(* IEC 61131-3 sources: PLC-IsaVODE/PLC-IsaVODE/samples/plc-programs (part 10) *)

(* ---- 683-FILE_PATH_SPLIT.ST ---- *)
TYPE
  oscat_STRING250             : STRING;
  oscat_STRING1             : STRING;
  oscat_STRING80             : STRING;
  oscat_STRING3             : STRING;
  oscat_NW_BUF_LONG  : ARRAY [0..4095] OF BYTE;
  PRINTF_DATA_250  	:  ARRAY [1..11]  OF oscat_STRING250;
  PRINTF_DATA_80 	:  ARRAY [1..11]  OF oscat_STRING80;
  LOG_250       	:  ARRAY [0..400] OF oscat_STRING250;
  LOG_80    		:  ARRAY [0..400] OF oscat_STRING80;
  LOG_OPTION		:  ARRAY [0..400] OF DWORD;

  us_LOG_CONTROL :
  STRUCT
    NEW_MSG              : oscat_STRING250;    (*W neue Nachricht f�r den Datenbuffer   *)
	NEW_MSG_OPTION 		 : DWORD;
    LEVEL                : BYTE;
	SIZE                 : INT;                (*R Anzahl der Strings im LOG_DATA       *)
	RESET                : BOOL;               (*W Nachrichtenbuffer l�schen            *)
    PRINTF               : PRINTF_DATA_250;    (*W Array PRINTF Parameter               *)
    MSG                  : LOG_250;            (*I Array Message                        *)
    MSG_OPTION           : LOG_OPTION;     	   (*I Array Message Option                 *)
	UPDATE_COUNT         : UINT;               (*R Updatez�hler                         *)
    IDX                  : INT;                (*R aktueller Nachrichten-Index          *)
	RING_MODE            : BOOL;               (*I Buffer�berlauf erkannt               *)
  END_STRUCT;

  us_LOG_CONTROL_80 :
  STRUCT
    NEW_MSG              : oscat_STRING80;     (*W neue Nachricht f�r den Datenbuffer   *)
	NEW_MSG_OPTION 		 : DWORD;
    LEVEL                : BYTE;
	SIZE                 : INT;                (*R Anzahl der Strings im LOG_DATA       *)
	RESET                : BOOL;               (*W Nachrichtenbuffer l�schen            *)
    PRINTF               : PRINTF_DATA_80;     (*W Array PRINTF Parameter               *)
    MSG                  : LOG_80;             (*I Array Message                        *)
    MSG_OPTION           : LOG_OPTION;     	   (*I Array Message Option                 *)
	UPDATE_COUNT         : UINT;               (*R Updatez�hler                         *)
    IDX                  : INT;                (*R aktueller Nachrichten-Index          *)
	RING_MODE            : BOOL;               (*I Buffer�berlauf erkannt               *)
  END_STRUCT;

  LINE_ARRAY 			: ARRAY [1..40] OF INT;

  us_LOG_VIEWPORT :
    STRUCT
     LINE_ARRAY          : LINE_ARRAY;
     COUNT               : INT;                (* Anzahl der sichtbaren Nachtrichten   *)
	 UPDATE_COUNT        : UINT;               (* Updatez�hler                         *)
     MOVE_TO_X           : INT;                (* Steuerung der Nachrichtenanzeige     *)
     UPDATE              : BOOL;               (* Daten wurden ge�ndert -> neuzeichnen *)
  END_STRUCT;

  oscat_FILE_SERVER_DATA : STRUCT
	FILE_OPEN	: BOOL;
    FILENAME 	: STRING;
    MODE	 	: BYTE;
    OFFSET   	: UDINT;
    FILE_SIZE   : UDINT;
    AUTO_CLOSE	: TIME;
    ERROR	 	: BYTE;
  END_STRUCT;

  oscat_FILE_PATH_DATA : STRUCT
	DRIVE : oscat_string3;
	DIRECTORY : oscat_string250;
	FILENAME : STRING;
  END_STRUCT;

  oscat_UNI_CIRCULAR_BUFFER_DATA : STRUCT
	D_MODE : INT;
	D_HEAD : WORD;
	D_STRING : oscat_string250;
	D_REAL : REAL;
	D_DWORD : DWORD;
	BUF_SIZE : INT;
	BUF_COUNT : INT;
	BUF_USED : USINT;
	BUF : oscat_NW_BUF_LONG;
	_GetStart : INT;
	_GetEnd : INT;
	_Last : INT;
	_First : INT;
  END_STRUCT;

  oscat_DLOG_DATA : STRUCT
	STORE_TYPE : BYTE;
	ADD_HEADER : BOOL;
	ADD_DATA : BOOL;
	ADD_DATA_REQ : BOOL;
	CLOCK_TRIG : BOOL;
	ID_MAX : USINT;
	DTI : UDINT;
	UCB : oscat_UNI_CIRCULAR_BUFFER_DATA;
	NEW_FILE : STRING;
	NEW_FILE_RTRIG : BOOL;
  END_STRUCT;

END_TYPE

FUNCTION_BLOCK FILE_PATH_SPLIT_Block

	VAR_INPUT
		FILENAME :	oscat_STRING250;
	END_VAR

	VAR_OUTPUT
		FILE_PATH_SPLIT :	BOOL;
	END_VAR

	VAR_IN_OUT
		X :	oscat_FILE_PATH_DATA;
	END_VAR

	VAR
		b :	INT;
		c :	INT;
		d :	oscat_STRING1;
		p1 :	INT;
		p2 :	INT;
	END_VAR

	X.DRIVE := '';
	X.DIRECTORY := '';
	X.FILENAME := '';
	p1 := 0;
	p2 := 0;
	c := LEN(FILENAME);
	IF c = 0 THEN
		FILE_PATH_SPLIT := FALSE;
		RETURN;
	END_IF;

	FOR b := 1 TO c DO
		d := MID(FILENAME, 1, b);
		IF EQ_STRING(d,':') THEN
			p1 := b;
		ELSIF EQ_STRING(d,'/') OR EQ_STRING(d,'\') THEN
			p2 := b;
		END_IF;
	END_FOR;

	IF p1 = 2 THEN
		X.DRIVE := LEFT(FILENAME,p1);
	END_IF;

	IF p2 > 0 AND p2 > p1 THEN
		X.DIRECTORY := MID(FILENAME,p2-p1,p1+1);
	END_IF;

	X.FILENAME := RIGHT(FILENAME,c - MAX (p1,p2));
	FILE_PATH_SPLIT := TRUE;

END_FUNCTION_BLOCK

PROGRAM program0
	VAR
		FILENAME :	oscat_STRING250;
		FILE_PATH_SPLIT :	BOOL;
		X :	oscat_FILE_PATH_DATA;

		func_block : FILE_PATH_SPLIT_Block;
	END_VAR
	func_block.FILENAME := FILENAME;
	func_block.X := X;

	func_block();
	FILE_PATH_SPLIT  := func_block.FILE_PATH_SPLIT;
	X  := func_block.X;
END_PROGRAM

CONFIGURATION Config0
	RESOURCE Res0 ON PLC
		TASK task0(INTERVAL := T#20ms,PRIORITY := 0);
		PROGRAM instance0 WITH task0 : program0;
	END_RESOURCE
END_CONFIGURATION

(* ---- 684-BLIND_SHADE.ST ---- *)
TYPE
  oscat_STRING5               : STRING;
  oscat_STRING30              : STRING;
END_TYPE

TYPE oscat_CALENDAR :
	STRUCT
		UTC : UDINT;				(* world time UTC *)
		LDT : UDINT;				(* local time *)
		LDATE : UDINT;				(* local date *)
		LTOD : UDINT;				(* local time of day *)
		YEAR : INT;					(* year of LDATE *)
		MONTH : INT;				(* month of LDATE *)
		DAY : INT;					(* day of LDATE *)
		WEEKDAY : INT;				(* weekday of LDATE *)
		OFFSET : INT;				(* Time Zone Offset for Local time in minutes *)
		DST_EN : BOOL;				(* daylight savings time enable *)
		DST_ON : BOOL;				(* true when daylight savings time os on *)
		NAME : oscat_string5;		(* name of time zone *)
		LANGUAGE : INT;			    (* language number pls see language setup *)
		LONGITUDE : REAL;			(* longitude of current location *)
		LATITUDE : REAL;			(* latitude of current location *)
		SUN_RISE : UDINT;			(* sun_rise for current location *)
		SUN_SET : UDINT;			(* sun_set for current location *)
		SUN_MIDDAY : UDINT;			(* worldtime when sun stands at south position *)
		SUN_HEIGTH : REAL;			(* suns heigth at midday, south position *)
		SUN_HOR : REAL;				(* sun angle horizontal 0 = north in degrees *)
		SUN_VER : REAL;				(* sun angle vertical above horizon in degrees *)
		NIGHT : BOOL;				(* true between sun_set and sun_rise *)
		HOLIDAY : BOOL;				(* true when holiday *)
		HOLY_NAME : oscat_string30;	(* name of holiday *)
		WORK_WEEK : INT;			(* current work week *)
	END_STRUCT;
END_TYPE

FUNCTION DT_TO_TOD2:UDINT
	VAR_INPUT
		IN :	UDINT;
	END_VAR

	DT_TO_TOD2 := (IN MOD UDINT#86400) * UDINT#1000;
END_FUNCTION

FUNCTION TIME_TO_UDINT2:UDINT
	VAR_INPUT
		X :	TIME;
	END_VAR

	TIME_TO_UDINT2 := DINT_TO_UDINT(TIME_TO_DINT(X));
END_FUNCTION

FUNCTION DEG : REAL
	VAR_INPUT
		RAD_IN : REAL;
	END_VAR

	DEG := MODR(57.29577951308232 * RAD_IN, 360.0);
END_FUNCTION

FUNCTION MODR : REAL
	VAR_INPUT
		IN : REAL;
		DIVI : REAL;
	END_VAR

	IF divi = 0.0 THEN
		MODR := 0.0;
	ELSE
		MODR := in - DINT_TO_REAL(FLOOR2(in / divi)) * divi;
	END_IF;
END_FUNCTION

FUNCTION FLOOR2 : DINT
	VAR_INPUT
		x : REAL;
	END_VAR

	FLOOR2 := REAL_TO_DINT(X);
	IF DINT_TO_REAL(FLOOR2) > X THEN
		FLOOR2 := FLOOR2 - DINT#1;
	END_IF;
END_FUNCTION

FUNCTION RAD:REAL

	VAR_INPUT
		DEG1 :	REAL;
	END_VAR

	RAD := MODR(0.0174532925199433 * DEG1 , 6.283185307179586476);

END_FUNCTION

FUNCTION TRUNC_UDINT2:UDINT
	VAR_INPUT
		IN :	REAL;
	END_VAR
	TRUNC_UDINT2 := DINT_TO_UDINT(TRUNC_DINT(IN));
END_FUNCTION

FUNCTION_BLOCK BLIND_SHADE_Block

	VAR_INPUT
		UP :	BOOL;
		DN :	BOOL;
		S_IN :	BYTE;
		PI :	BYTE;
		AI :	BYTE;
		ENABLE :	BOOL;
		SUN :	BOOL;
		SUNRISE_OFFSET :	TIME := T#1h;
		SUNSET_PRESET :	TIME := T#1h;
		DIRECTION :	REAL := 180.0;
		ANGLE_OFFSET :	REAL := 80.0;
		SLAT_WIDTH :	REAL := 80.0;
		SLAT_SPACING :	REAL := 60.0;
		SHADE_DELAY :	TIME := T#60s;
		SHADE_POS :	BYTE;
	END_VAR

	VAR_OUTPUT
		QU :	BOOL;
		QD :	BOOL;
		STATUS :	BYTE;
		PO :	BYTE;
		AO :	BYTE;
	END_VAR

	VAR_IN_OUT
		CX :	oscat_CALENDAR;
	END_VAR

	VAR
		angle :	REAL;
		sun_delay :	TOF;
	END_VAR

	sun_delay(IN := sun, PT := shade_delay);

	IF UP AND DN AND enable AND sun_delay.Q AND cx.SUN_HOR > direction - angle_offset AND cx.SUN_HOR < direction + angle_offset AND
		DT_TO_TOD2(cx.UTC) > cx.SUN_RISE + TIME_TO_UDINT2(sunrise_offset) AND DT_TO_TOD2(cx.UTC) < cx.SUN_SET - TIME_TO_UDINT2(sunset_preset) THEN
		status := BYTE#151;
		QU := UP;
		QD := DN;
		po := shade_pos;
		angle := DEG(ATAN(slat_spacing / slat_width));
		IF cx.SUN_VER > 0.0 AND cx.SUN_VER < angle THEN
			angle := cx.SUN_VER + DEG(ACOS(COS(RAD(cx.SUN_VER))*slat_spacing / Slat_width));
			ao := INT_TO_BYTE(LIMIT(0,UDINT_TO_INT(TRUNC_UDINT2(angle * 2.833333333)), 255));
		ELSE
			ao := BYTE#255;
		END_IF;
	ELSE
		QU := UP;
		QD := DN;
		po := pi;
		ao := ai;
		status := S_IN;
	END_IF;

END_FUNCTION_BLOCK

PROGRAM program0
	VAR
		UP :	BOOL;
		DN :	BOOL;
		S_IN :	BYTE;
		PI :	BYTE;
		AI :	BYTE;
		ENABLE :	BOOL;
		SUN :	BOOL;
		SUNRISE_OFFSET :	TIME := T#1h;
		SUNSET_PRESET :	TIME := T#1h;
		DIRECTION :	REAL := 180.0;
		ANGLE_OFFSET :	REAL := 80.0;
		SLAT_WIDTH :	REAL := 80.0;
		SLAT_SPACING :	REAL := 60.0;
		SHADE_DELAY :	TIME := T#60s;
		SHADE_POS :	BYTE;
		CX :	oscat_CALENDAR;

		func_block : BLIND_SHADE_Block;
	END_VAR
	func_block.UP := UP;
	func_block.DN := DN;
	func_block.S_IN := S_IN ;
	func_block.PI    := PI    ;
	func_block.AI    := AI    ;
	func_block.ENABLE := ENABLE;
	func_block.SUN := SUN;
	func_block.SUNRISE_OFFSET := SUNRISE_OFFSET;
	func_block.SUNSET_PRESET := SUNSET_PRESET ;
	func_block.DIRECTION := DIRECTION ;
	func_block.ANGLE_OFFSET    := ANGLE_OFFSET    ;
	func_block.SLAT_WIDTH := SLAT_WIDTH;
	func_block.SLAT_SPACING := SLAT_SPACING;
	func_block.SHADE_DELAY := SHADE_DELAY ;
	func_block.CX := CX ;

	func_block();
	CX  := func_block.CX;
END_PROGRAM

CONFIGURATION Config0
	RESOURCE Res0 ON PLC
		TASK task0(INTERVAL := T#20ms,PRIORITY := 0);
		PROGRAM instance0 WITH task0 : program0;
	END_RESOURCE
END_CONFIGURATION

(* ---- 686-_ARRAY_SHUFFLE.ST ---- *)
TYPE
	oscat_pt_ARRAY: ARRAY [1..100] OF REAL;
END_TYPE

FUNCTION D_TRUNC : DINT
  VAR_INPUT
    x : REAL;
  END_VAR

  D_TRUNC := REAL_TO_DINT(X);
  IF X > 0.0 THEN
  	IF DINT_TO_REAL(D_TRUNC) > X THEN D_TRUNC := D_TRUNC - DINT#1; END_IF;
  ELSE
  	IF DINT_TO_REAL(D_TRUNC) < X THEN D_TRUNC := D_TRUNC + DINT#1; END_IF;
  END_IF;
END_FUNCTION

FUNCTION BIT_COUNT:INT
	VAR_INPUT
		IN :	DWORD;
	END_VAR

	VAR
		in_temp :	DWORD;
	END_VAR

	in_temp := IN;
	WHILE in_temp > DWORD#0 DO
		IF (in_temp AND DWORD#16#00000001) > DWORD#0 THEN Bit_Count := Bit_Count +1; END_IF;
		in_temp := SHR(in_temp,1);
	END_WHILE;
END_FUNCTION

FUNCTION FRACT:REAL
	VAR_INPUT
		X :	REAL;
	END_VAR

	IF ABS(x) < 2.0E9 THEN
		FRACT := x - DINT_TO_REAL(D_TRUNC(x));
	ELSE
		FRACT := 0.0;
	END_IF;
END_FUNCTION

FUNCTION_BLOCK T_PLC_MS_block
	VAR_OUTPUT
		T_PLC_MS :	UDINT;
	END_VAR

	VAR_EXTERNAL
		PLC_TICKS_PER_SEC :	INT;
		PLC_SYS_TICK_CNT :	DINT;
	END_VAR

	VAR
		debug :	BOOL;(*Debug-Mode ON / OFF*)
		N :	INT;(*Debug-Faktor*)
		Offset :	UDINT;(*Debug-Offset*)
		temp :	DWORD := DWORD#1;(*Debug-Offset*)
		mode :	BOOL;(*modus*)
		faktor :	UDINT;(*Systemtakt-Faktor*)
		init :	BOOL;
		v_plc_ticks_per_sec :	UDINT;
		base :	UDINT := UDINT#1000;
	END_VAR

	IF init = FALSE THEN
		v_plc_ticks_per_sec := INT_TO_UDINT(PLC_TICKS_PER_SEC);
		IF v_plc_ticks_per_sec = UDINT#1024 THEN
			faktor := UDINT#1;
			mode := FALSE;
		ELSIF v_plc_ticks_per_sec > UDINT#0 THEN
			IF v_plc_ticks_per_sec <= base THEN
				faktor := base / v_plc_ticks_per_sec;
				mode := FALSE;
			ELSE
				faktor := v_plc_ticks_per_sec / base;
				mode := TRUE;
			END_IF;
		ELSE
			faktor := UDINT#1;
		END_IF;
		init := TRUE;
	END_IF;

	IF mode THEN
		T_PLC_MS := DINT_TO_UDINT(PLC_SYS_TICK_CNT) / faktor;
	ELSE
		T_PLC_MS := DINT_TO_UDINT(PLC_SYS_TICK_CNT) * faktor;
	END_IF;

	IF debug THEN
		T_PLC_MS := (DWORD_TO_UDINT(SHL(UDINT_TO_DWORD(T_PLC_MS),N) OR SHL(temp,N)) - UDINT#1) + Offset;
	END_IF;
END_FUNCTION_BLOCK

FUNCTION BIT_LOAD_DW:DWORD

	VAR_INPUT
		IN :	DWORD;
		VAL :	BOOL;
		POS :	INT;
	END_VAR

	IF val THEN
		BIT_LOAD_DW := in OR SHL(DWORD#1,pos);
	ELSE
		BIT_LOAD_DW := in AND (NOT SHL(DWORD#1,pos));
	END_IF;
END_FUNCTION

FUNCTION BIT_OF_DWORD : BOOL
  VAR_INPUT
    IN : DWORD;
    N : INT;
  END_VAR

  BIT_OF_DWORD := (SHR(in,N) AND 16#00000001) > 0;
  (* from OSCAT library; www.oscat.de  *)
END_FUNCTION

FUNCTION _INT_TO_UDINT:UDINT
	VAR_INPUT
		IN :	INT;
	END_VAR

	_INT_TO_UDINT := DINT_TO_UDINT(INT_TO_DINT(IN));
END_FUNCTION

FUNCTION _DWORD_TO_REAL:REAL
	VAR_INPUT
		IN :	DWORD;
	END_VAR

	_DWORD_TO_REAL := UDINT_TO_REAL(DWORD_TO_UDINT(IN));

END_FUNCTION

FUNCTION_BLOCK RDM_block
	VAR_INPUT
		LAST :	REAL;
	END_VAR
	VAR_OUTPUT
		RDM :	REAL;
	END_VAR
	VAR
		T_PLC_MS :	T_PLC_MS_block;
		tn :	DWORD;
		tc :	INT;
	END_VAR
	T_PLC_MS();
	tn := UDINT_TO_DWORD(T_PLC_MS.T_PLC_MS);
	tc := Bit_Count(tn);

	tn:=BIT_LOAD_DW(tn,BIT_OF_DWORD(tn,2),31); (* tn.31 := tn.2; *)
	tn:=BIT_LOAD_DW(tn,BIT_OF_DWORD(tn,5),30); (* tn.30 := tn.5; *)
	tn:=BIT_LOAD_DW(tn,BIT_OF_DWORD(tn,4),29); (* tn.29 := tn.4; *)
	tn:=BIT_LOAD_DW(tn,BIT_OF_DWORD(tn,1),28); (* tn.28 := tn.1; *)
	tn:=BIT_LOAD_DW(tn,BIT_OF_DWORD(tn,0),27); (* tn.27 := tn.0; *)
	tn:=BIT_LOAD_DW(tn,BIT_OF_DWORD(tn,7),26); (* tn.26 := tn.7; *)
	tn:=BIT_LOAD_DW(tn,BIT_OF_DWORD(tn,6),25); (* tn.25 := tn.6; *)
	tn:=BIT_LOAD_DW(tn,BIT_OF_DWORD(tn,3),24); (* tn.24 := tn.3; *)

	tn := ROL(tn,Bit_Count(tn)) OR DWORD#16#80000001;
	tn := UDINT_TO_DWORD(DWORD_TO_UDINT(tn) MOD UDINT#71474513 + _INT_TO_UDINT(tc) + UDINT#77);
	RDM := fract(_DWORD_TO_REAL(tn) / 10000000.0 * (2.71828182845904523536028747135266249 - LIMIT_REAL(0.0,last,1.0)));
END_FUNCTION_BLOCK

FUNCTION_BLOCK RDM22
	VAR_INPUT
		LAST :	INT;
		LOW :	INT;
		HIGH :	INT;
	END_VAR

	VAR_OUTPUT
		RDM2 :	INT;
	END_VAR

	VAR
		rdm :	RDM_block;
	END_VAR

	rdm(last:=fract(INT_TO_REAL(last) * 3.14159265358979323846264338327950288));
	RDM2 := TRUNC(rdm.RDM * INT_TO_REAL(high - low + 1)) + low;
END_FUNCTION_BLOCK

FUNCTION_BLOCK _ARRAY_SHUFFLE2
	VAR_IN_OUT
		PT :	oscat_pt_ARRAY;
	END_VAR

	VAR_INPUT
		SIZE :	UINT;
	END_VAR

	VAR_OUTPUT
		_ARRAY_SHUFFLE :	BOOL;
	END_VAR
	VAR
		temp :	REAL;
		pos :	INT;
		i :	INT;
		stop :	INT;
		rdm2 :	rdm22;
	END_VAR

	stop :=LIMIT_INT(1,UINT_TO_INT(size),1000);
	FOR i := 1 TO stop DO
			rdm2(last:=i+pos,low:=1,high:=stop);
			pos := rdm2.rdm2;
			(* swap elements *)
			temp := pt[i];
			pt[i] := pt[pos];
			pt[pos] := temp;
	END_FOR;

	_ARRAY_SHUFFLE := TRUE;
END_FUNCTION_BLOCK

PROGRAM program0
  VAR
    LocalVar0 : oscat_pt_ARRAY;
    LocalVar1 : UINT;
	LocalOUT  : BOOL;
	func_block : _ARRAY_SHUFFLE2;
  END_VAR
	func_block.pt := LocalVar0;
	func_block.size := LocalVar1;
	func_block();
	LocalOUT := func_block._ARRAY_SHUFFLE;

END_PROGRAM

CONFIGURATION Config0
	VAR_GLOBAL
		PLC_TICKS_PER_SEC :	INT;
		PLC_SYS_TICK_CNT :	DINT;
	END_VAR
  RESOURCE Res0 ON PLC
    TASK task0(INTERVAL := T#20ms,PRIORITY := 0);
    PROGRAM instance0 WITH task0 : program0;
  END_RESOURCE
END_CONFIGURATION

(* ---- 687-TN_INPUT_SELECT_TEXT.ST ---- *)
TYPE
  bya_TN_CHAR:       	ARRAY [0..1919] OF BYTE;
  bya_TN_BACKUP:     	ARRAY [0..1919] OF BYTE;
  bya_TN_COLOR:      	ARRAY [0..1919] OF BYTE;
  bya_TN_Line_Update:	ARRAY [0..23]   OF BOOL;

  us_TN_SCREEN :
  STRUCT
		bya_CHAR:			bya_TN_CHAR;
		bya_COLOR:			bya_TN_COLOR;
		bya_BACKUP:			bya_TN_BACKUP;
		bya_Line_Update:	bya_TN_Line_Update;

		by_Input_Exten_Code:    BYTE;
		by_Input_ASCII_Code:    BYTE;
		bo_Input_ASCII_IsNum:   BOOL;
		in_Page_Number:        	INT;
		in_Cursor_X:           	INT;
		in_Cursor_Y:           	INT;
		in_EOS_Offset:         	INT;
		by_Clear_Screen_Attr:  	BYTE;
		bo_Clear_Screen:       	BOOL;
		bo_Modal_Dialog:       	BOOL;
		bo_Menue_Bar_Dialog:   	BOOL;

  END_STRUCT;
END_TYPE

FUNCTION_BLOCK TN_INPUT_SELECT_TEXT_Block

  VAR
    in_count :	INT;
    by_Attr :	BYTE;
    st_String :	STRING;
  END_VAR

  VAR
    FB_FIX :	FIX;
    FB_TN_SC_WRITE :	TN_SC_WRITE;
    ELEMENT_COUNT :	ELEMENT_COUNT;
    ELEMENT_GET :	ELEMENT_GET;
  END_VAR

  VAR_IN_OUT
    Xus_TN_SCREEN :	us_TN_SCREEN;
    Xus_TN_INPUT_CONTROL_DATA :	us_TN_INPUT_CONTROL_DATA;
  END_VAR

  IF Xus_TN_INPUT_CONTROL_DATA.bo_Focus = TRUE THEN

    IF Xus_TN_INPUT_CONTROL_DATA.by_Input_ASCII_Code = BYTE#32 THEN
      Xus_TN_INPUT_CONTROL_DATA.in_selected := Xus_TN_INPUT_CONTROL_DATA.in_selected + INT#01;
      Xus_TN_INPUT_CONTROL_DATA.bo_Update_Input := TRUE;
    END_IF;

    IF Xus_TN_INPUT_CONTROL_DATA.by_Input_Exten_Code = BYTE#13 THEN
      Xus_TN_INPUT_CONTROL_DATA.bo_Input_Entered := TRUE;
    END_IF;

  END_IF;

  IF (Xus_TN_INPUT_CONTROL_DATA.bo_Update_Input = TRUE) OR (Xus_TN_INPUT_CONTROL_DATA.bo_Update_All = TRUE) THEN

    IF Xus_TN_INPUT_CONTROL_DATA.bo_Update_All = TRUE THEN

      IF (Xus_TN_INPUT_CONTROL_DATA.in_Title_X_Offset = INT#00) AND (Xus_TN_INPUT_CONTROL_DATA.in_Title_Y_Offset = INT#00) THEN

        FB_TN_SC_WRITE.Iin_Y := Xus_TN_INPUT_CONTROL_DATA.in_Y;
        FB_TN_SC_WRITE.Iin_X := Xus_TN_INPUT_CONTROL_DATA.in_X - LEN(Xus_TN_INPUT_CONTROL_DATA.st_Title_String);

      ELSE
        FB_TN_SC_WRITE.Iin_Y := Xus_TN_INPUT_CONTROL_DATA.in_Y + Xus_TN_INPUT_CONTROL_DATA.in_Title_Y_Offset;
        FB_TN_SC_WRITE.Iin_X := Xus_TN_INPUT_CONTROL_DATA.in_X + Xus_TN_INPUT_CONTROL_DATA.in_Title_X_Offset;

      END_IF;

      FB_TN_SC_WRITE.Iby_ATTR      := Xus_TN_INPUT_CONTROL_DATA.by_Title_Attr;
      FB_TN_SC_WRITE.Ist_STRING    := Xus_TN_INPUT_CONTROL_DATA.st_Title_String;
      FB_TN_SC_WRITE.Xus_TN_SCREEN := Xus_TN_SCREEN;
      FB_TN_SC_WRITE();
      Xus_TN_SCREEN := FB_TN_SC_WRITE.Xus_TN_SCREEN;

    END_IF;

    ELEMENT_COUNT(ELEMENT:=Xus_TN_INPUT_CONTROL_DATA.st_Input_Data,SEP:=BYTE#35);
    Xus_TN_INPUT_CONTROL_DATA.st_Input_Data:=ELEMENT_COUNT.ELEMENT;
    in_count:=ELEMENT_COUNT.ELEMENT_COUNT;

    IF in_Count > INT#00 THEN

      IF Xus_TN_INPUT_CONTROL_DATA.in_selected < INT#1 THEN
        Xus_TN_INPUT_CONTROL_DATA.in_selected := INT#01;
      END_IF;

      IF Xus_TN_INPUT_CONTROL_DATA.in_selected > in_count THEN
        Xus_TN_INPUT_CONTROL_DATA.in_selected := INT#01;
      END_IF;

      ELEMENT_GET(ELEMENT:=Xus_TN_INPUT_CONTROL_DATA.st_Input_Data,SEP:=BYTE#35,POS:=Xus_TN_INPUT_CONTROL_DATA.in_selected-1);
      Xus_TN_INPUT_CONTROL_DATA.st_Input_Data := ELEMENT_GET.ELEMENT;
      st_String:=ELEMENT_GET.ELEMENT_GET;

      FB_FIX.str:=st_String;
    FB_FIX.L:=LEN(Xus_TN_INPUT_CONTROL_DATA.st_Input_Mask);
    FB_FIX.C:=BYTE#32;
    FB_FIX.M:=Xus_TN_INPUT_CONTROL_DATA.in_Input_Option;
      FB_FIX();
      st_String:=FB_FIX.FIX;

      Xus_TN_INPUT_CONTROL_DATA.st_Input_String := st_String;

      IF Xus_TN_INPUT_CONTROL_DATA.bo_Focus = TRUE THEN
        by_Attr := Xus_TN_INPUT_CONTROL_DATA.by_Attr_mF;
      ELSE
        by_Attr := Xus_TN_INPUT_CONTROL_DATA.by_Attr_oF;
      END_IF;

      FB_TN_SC_WRITE.Iin_Y         := Xus_TN_INPUT_CONTROL_DATA.in_Y;
      FB_TN_SC_WRITE.Iin_X         := Xus_TN_INPUT_CONTROL_DATA.in_X;
      FB_TN_SC_WRITE.Iby_ATTR      := by_Attr;
      FB_TN_SC_WRITE.Ist_STRING    := st_String;
      FB_TN_SC_WRITE.Xus_TN_SCREEN := Xus_TN_SCREEN;
      FB_TN_SC_WRITE();
      Xus_TN_SCREEN := FB_TN_SC_WRITE.Xus_TN_SCREEN;

    END_IF;

    Xus_TN_INPUT_CONTROL_DATA.in_Cursor_Y := Xus_TN_INPUT_CONTROL_DATA.in_Y;
    Xus_TN_INPUT_CONTROL_DATA.in_Cursor_X := Xus_TN_INPUT_CONTROL_DATA.in_X;

    Xus_TN_INPUT_CONTROL_DATA.bo_Update_All   := FALSE;
    Xus_TN_INPUT_CONTROL_DATA.bo_Update_Input := FALSE;

  END_IF;

END_FUNCTION_BLOCK

PROGRAM program0
	VAR
		Xus_TN_SCREEN :	us_TN_SCREEN;
    Xus_TN_INPUT_CONTROL_DATA :	us_TN_INPUT_CONTROL_DATA;

		func_block : TN_INPUT_SELECT_TEXT_Block;
	END_VAR
	func_block.Xus_TN_INPUT_CONTROL_DATA := Xus_TN_INPUT_CONTROL_DATA;
	func_block.Xus_TN_SCREEN := Xus_TN_SCREEN;

	func_block();
  Xus_TN_INPUT_CONTROL_DATA  := func_block.Xus_TN_INPUT_CONTROL_DATA;
	Xus_TN_SCREEN  := func_block.Xus_TN_SCREEN;
END_PROGRAM

CONFIGURATION Config0
	RESOURCE Res0 ON PLC
		TASK task0(INTERVAL := T#20ms,PRIORITY := 0);
		PROGRAM instance0 WITH task0 : program0;
	END_RESOURCE
END_CONFIGURATION

(* ---- 688-SEQUENCE_4.ST ---- *)
FUNCTION UDINT_TO_TIME2:TIME

	VAR_INPUT
		IN :	UDINT;
	END_VAR

	UDINT_TO_TIME2 := DINT_TO_TIME(UDINT_TO_DINT(IN));

END_FUNCTION

FUNCTION_BLOCK T_PLC_MS_block
	VAR_OUTPUT
		T_PLC_MS :	UDINT;
	END_VAR

	VAR_EXTERNAL
		PLC_TICKS_PER_SEC :	INT;
		PLC_SYS_TICK_CNT :	DINT;
	END_VAR

	VAR
		debug :	BOOL;
		N :	INT;
		Offset :	UDINT;
		temp :	DWORD := DWORD#1;
		mode :	BOOL;
		faktor :	UDINT;
		init :	BOOL;
		v_plc_ticks_per_sec :	UDINT;
		base :	UDINT := UDINT#1000;
	END_VAR

	IF init = FALSE THEN
		v_plc_ticks_per_sec := INT_TO_UDINT(PLC_TICKS_PER_SEC);
		IF v_plc_ticks_per_sec = UDINT#1024 THEN
			faktor := UDINT#1;
			mode := FALSE;
		ELSIF v_plc_ticks_per_sec > UDINT#0 THEN
			IF v_plc_ticks_per_sec <= base THEN
				faktor := base / v_plc_ticks_per_sec;
				mode := FALSE;
			ELSE
				faktor := v_plc_ticks_per_sec / base;
				mode := TRUE;
			END_IF;
		ELSE
			faktor := UDINT#1;
		END_IF;
		init := TRUE;
	END_IF;

	IF mode THEN
		T_PLC_MS := DINT_TO_UDINT(PLC_SYS_TICK_CNT) / faktor;
	ELSE
		T_PLC_MS := DINT_TO_UDINT(PLC_SYS_TICK_CNT) * faktor;
	END_IF;

	IF debug THEN
		T_PLC_MS := (DWORD_TO_UDINT(SHL(UDINT_TO_DWORD(T_PLC_MS),N) OR SHL(temp,N)) - UDINT#1) + Offset;
	END_IF;

END_FUNCTION_BLOCK

FUNCTION_BLOCK SEQUENCE_4_Block

	VAR_INPUT
		IN0 :	BOOL := TRUE;
		IN1 :	BOOL := TRUE;
		IN2 :	BOOL := TRUE;
		IN3 :	BOOL := TRUE;
		START :	BOOL;
		RST :	BOOL;
		WAIT0 :	TIME;
		DELAY0 :	TIME;
		WAIT1 :	TIME;
		DELAY1 :	TIME;
		WAIT2 :	TIME;
		DELAY2 :	TIME;
		WAIT3 :	TIME;
		DELAY3 :	TIME;
		STOP_ON_ERROR :	BOOL;
	END_VAR

	VAR_OUTPUT
		Q0 :	BOOL;
		Q1 :	BOOL;
		Q2 :	BOOL;
		Q3 :	BOOL;
		QX :	BOOL;
		RUN :	BOOL;
		_STEP :	INT := -1;
		STATUS :	BYTE;
	END_VAR

	VAR
		last :	TIME;
		edge :	BOOL;
		tx :	TIME;
		init :	BOOL;
		T_PLC_MS :	T_PLC_MS_Block;
	END_VAR

	T_PLC_MS();
	tx:= UDINT_TO_TIME(T_PLC_MS.T_PLC_MS);

	IF NOT init THEN
		last := tx;
		init := TRUE;
		status := BYTE#110;
	END_IF;

	IF rst THEN
		_step := -1;
		Q0 := FALSE;
		Q1 := FALSE;
		Q2 := FALSE;
		Q3 := FALSE;
		status := BYTE#110;
		run := FALSE;

	ELSIF start AND NOT edge THEN
		_step := 0;
		last := tx;
		status := BYTE#111;
		Q0 := FALSE;
		Q1 := FALSE;
		Q2 := FALSE;
		Q3 := FALSE;
		run := TRUE;
	END_IF;
	edge := start;

	IF status > BYTE#0 AND status < BYTE#100 AND stop_on_error THEN RETURN; END_IF;

	IF run AND _step = 0 THEN
		IF NOT q0 AND in0 AND tx - last <= wait0 THEN
			Q0 := TRUE;
			last := tx;
		ELSIF NOT q0 AND tx - last > wait0 THEN
			status := BYTE#1;
			run := FALSE;
		ELSIF q0 AND tx - last >= delay0 THEN
			_step := 1;
			last := tx;
		END_IF;
	END_IF;
	IF run AND _step = 1 THEN
		IF NOT q1 AND in1 AND tx - last <= wait1 THEN
			Q0 := FALSE;
			Q1 := TRUE;
			last := tx;
		ELSIF NOT q1 AND Tx - last > wait1 THEN
			status := BYTE#2;
			q0 := FALSE;
			run := FALSE;
		ELSIF q1 AND tx - last >= delay1 THEN
			_step := 2;
			last := tx;
		END_IF;
	END_IF;
	IF run AND _step = 2 THEN
		IF NOT q2 AND in2 AND tx - last <= wait2 THEN
			Q1 := FALSE;
			Q2 := TRUE;
			last := tx;
		ELSIF NOT q2 AND Tx - last > wait2 THEN
			status := BYTE#3;
			q1 := FALSE;
			run := FALSE;
		ELSIF q2 AND tx - last >= delay2 THEN
			_step := 3;
			last := tx;
		END_IF;
	END_IF;
	IF run AND _step = 3 THEN
		IF NOT q3 AND in3 AND tx - last <= wait3 THEN
			Q2 := FALSE;
			Q3 := TRUE;
			last := tx;
		ELSIF NOT q3 AND Tx - last > wait3 THEN
			status := BYTE#4;
			q2 := FALSE;
			run := FALSE;
		ELSIF q3 AND tx - last >= delay3 THEN
			_step := -1;
			q3 := FALSE;
			run := FALSE;
			status := BYTE#110;
		END_IF;
	END_IF;
	QX := q0 OR q1 OR q2 OR q3;

END_FUNCTION_BLOCK

PROGRAM program0

	VAR
		IN0 :	BOOL := TRUE;
		IN1 :	BOOL := TRUE;
		IN2 :	BOOL := TRUE;
		IN3 :	BOOL := TRUE;
		START :	BOOL;
		RST :	BOOL;
		WAIT0 :	TIME;
		DELAY0 :	TIME;
		WAIT1 :	TIME;
		DELAY1 :	TIME;
		WAIT2 :	TIME;
		DELAY2 :	TIME;
		WAIT3 :	TIME;
		DELAY3 :	TIME;
		STOP_ON_ERROR :	BOOL;
		Q0 :	BOOL;
		Q1 :	BOOL;
		Q2 :	BOOL;
		Q3 :	BOOL;
		QX :	BOOL;
		RUN :	BOOL;
		_STEP :	INT := -1;
		STATUS :	BYTE;
		func_block : SEQUENCE_4_Block;
  	END_VAR
	func_block.IN0  :=IN0;
	func_block.IN1  :=IN1;
	func_block.IN2  :=IN2;
	func_block.IN3  :=IN3;
	func_block.START  :=START;
	func_block.RST  :=RST;
	func_block.WAIT0  :=WAIT0;
	func_block.DELAY0  :=DELAY0;
	func_block.WAIT1:=WAIT1;
	func_block.DELAY1:=DELAY1;
	func_block.WAIT2  :=WAIT2;
	func_block.DELAY2  :=DELAY2;
	func_block.WAIT3  :=WAIT3;
	func_block.DELAY3  :=DELAY3;
	func_block.DELAY1:=DELAY1;
	func_block.WAIT2  :=WAIT2;
	func_block.DELAY2  :=DELAY2;
	func_block.WAIT3  :=WAIT3;
	func_block.DELAY3  :=DELAY3;
	func_block.STOP_ON_ERROR  :=STOP_ON_ERROR;
	func_block();
	Q0 := func_block.Q0;
	Q1 := func_block.Q1;
	Q2 := func_block.Q2;
	Q3 := func_block.Q3;
	QX := func_block.QX;
	RUN := func_block.RUN;
	_STEP := func_block._STEP;
	STATUS := func_block.STATUS;

END_PROGRAM

CONFIGURATION Config0

	VAR_GLOBAL
		PLC_TICKS_PER_SEC :	INT;
		PLC_SYS_TICK_CNT :	DINT;
	END_VAR

	RESOURCE Res0 ON PLC
		TASK task0(INTERVAL := T#20ms,PRIORITY := 0);
		PROGRAM instance0 WITH task0 : program0;
	END_RESOURCE

END_CONFIGURATION

(* ---- 689-TN_SC_LINE.ST ---- *)
TYPE
  bya_TN_CHAR:       	ARRAY [0..1919] OF BYTE;
  bya_TN_BACKUP:     	ARRAY [0..1919] OF BYTE;
  bya_TN_COLOR:      	ARRAY [0..1919] OF BYTE;
  bya_TN_Line_Update:	ARRAY [0..23]   OF BOOL;

  us_TN_SCREEN :
  STRUCT
		bya_CHAR:			bya_TN_CHAR;
		bya_COLOR:			bya_TN_COLOR;
		bya_BACKUP:			bya_TN_BACKUP;
		bya_Line_Update:	bya_TN_Line_Update;

		by_Input_Exten_Code:    BYTE;
		by_Input_ASCII_Code:    BYTE;
		bo_Input_ASCII_IsNum:   BOOL;
		in_Page_Number:        	INT;                (* aktive Seiten-Nr.              *)
		in_Cursor_X:           	INT;                (* Cursor X-Position              *)
		in_Cursor_Y:           	INT;                (* Cursor Y-Position              *)
		in_EOS_Offset:         	INT;                (* End of String Offset           *)
		by_Clear_Screen_Attr:  	BYTE;               (* Clear-Screen Attr              *)
		bo_Clear_Screen:       	BOOL;               (* Clear-Screen ausl�sen          *)
		bo_Modal_Dialog:       	BOOL;               (* Modaler Dialog ist aktiv       *)
		bo_Menue_Bar_Dialog:   	BOOL;               (* Menue Dialog ist aktiv         *)

  END_STRUCT;
END_TYPE

FUNCTION TN_SC_XY2_ERROR:BOOL

	VAR_INPUT
		X1 :	INT;
		Y1 :	INT;
		X2 :	INT;
		Y2 :	INT;
	END_VAR

	TN_SC_XY2_ERROR := Y1 < 0 OR X1 < 0 OR Y2 < 0 OR X2 < 0 OR Y1 > 23 OR X1 > 79 OR Y2 > 23 OR X2 > 79;

END_FUNCTION

FUNCTION_BLOCK TN_SC_LINE_Block

  VAR
    by_Connect_Left_Char :	BYTE;
    by_Connect_Right_Char :	BYTE;
    by_Connect_Top_Char :	BYTE;
    by_Connect_Bottom_Char :	BYTE;
    by_Connect_Cruz_Char :	BYTE;
    by_Vertikal_Line_Char :	BYTE;
    by_Horzontal_Line_Char :	BYTE;
    by_old_Char :	BYTE;
    in_Offset_1 :	INT;
    in_ROW_Index :	INT;
    in_COL_Index :	INT;
    by_Char :	BYTE;
  END_VAR

  VAR_INPUT
    Iin_X1 :	INT;
    Iin_Y1 :	INT;
    Iin_X2 :	INT;
    Iin_Y2 :	INT;
    Iby_ATTR :	BYTE;
    Iby_BORDER :	BYTE;
  END_VAR

  VAR_IN_OUT
    Xus_TN_SCREEN :	us_TN_SCREEN;
  END_VAR

  IF TN_SC_XY2_ERROR(Iin_X1,Iin_Y1,Iin_X2,Iin_Y2) THEN RETURN; END_IF;

  IF Iby_Border = BYTE#01 THEN

    by_Connect_Top_Char    := BYTE#16#C2;
    by_Connect_Bottom_Char := BYTE#16#C1;
    by_Connect_Left_Char   := BYTE#16#C3;
    by_Connect_Right_Char  := BYTE#16#B4;
    by_Horzontal_Line_Char := BYTE#16#C4;
    by_Vertikal_Line_Char  := BYTE#16#B3;
    by_Connect_Cruz_Char   := BYTE#16#C5;

  ELSIF Iby_Border = BYTE#02 THEN

    by_Connect_Top_Char    := BYTE#16#CB;
    by_Connect_Bottom_Char := BYTE#16#CA;
    by_Connect_Left_Char   := BYTE#16#CC;
    by_Connect_Right_Char  := BYTE#16#B9;
    by_Horzontal_Line_Char := BYTE#16#CD;
    by_Vertikal_Line_Char  := BYTE#16#BA;
    by_Connect_Cruz_Char   := BYTE#16#CE;

  ELSE
    by_Connect_Top_Char    := Iby_Border;
    by_Connect_Bottom_Char := Iby_Border;
    by_Connect_Left_Char   := Iby_Border;
    by_Connect_Right_Char  := Iby_Border;
    by_Horzontal_Line_Char := Iby_Border;
    by_Vertikal_Line_Char  := Iby_Border;
    by_Connect_Cruz_Char   := Iby_Border;

  END_IF;

  IF Iin_X1 = Iin_X2 THEN

    in_Offset_1 := (Iin_Y1 * 80) + Iin_X1;

    FOR in_ROW_Index := Iin_Y1 TO Iin_Y2 DO

      by_old_Char := Xus_TN_SCREEN.bya_CHAR[in_Offset_1];

      by_Char := by_Vertikal_Line_Char;

      IF by_old_Char = by_Horzontal_Line_Char THEN

        IF in_ROW_Index = Iin_Y1 THEN
          by_Char := by_Connect_Top_Char;

        ELSIF in_ROW_Index = Iin_Y2 THEN
          by_Char := by_Connect_Bottom_Char;

        ELSE
          by_Char := by_Connect_Cruz_Char;
        END_IF;

      END_IF;

      Xus_TN_SCREEN.bya_Line_Update[in_ROW_Index] := TRUE;

      Xus_TN_SCREEN.bya_CHAR[in_Offset_1]  := by_Char;
      Xus_TN_SCREEN.bya_COLOR[in_Offset_1] := Iby_Attr;

      in_Offset_1 := in_Offset_1 + 80;

    END_FOR;

  ELSIF Iin_Y1 = Iin_Y2 THEN

    Xus_TN_SCREEN.bya_Line_Update[Iin_Y1] := TRUE;

    in_Offset_1 := (Iin_Y1 * 80) + Iin_X1;

    FOR in_COL_Index := Iin_X1 TO Iin_X2 DO

      by_old_Char := Xus_TN_SCREEN.bya_CHAR[in_Offset_1];

      by_Char := by_Horzontal_Line_Char;

      IF by_old_Char = by_Vertikal_Line_Char THEN

        IF in_COL_Index = Iin_X1 THEN
          by_Char := by_Connect_Left_Char;

        ELSIF in_COL_Index = Iin_X2 THEN
          by_Char := by_Connect_Right_Char;

        ELSE
          by_Char := by_Connect_Cruz_Char;
        END_IF;

      END_IF;

      Xus_TN_SCREEN.bya_CHAR[in_Offset_1]  := by_Char;
      Xus_TN_SCREEN.bya_COLOR[in_Offset_1] := Iby_Attr;

      in_Offset_1 := in_Offset_1 + 1;

    END_FOR;
  END_IF;

END_FUNCTION_BLOCK

PROGRAM program0
	VAR
    Iin_X1 :	INT;
    Iin_Y1 :	INT;
    Iin_X2 :	INT;
    Iin_Y2 :	INT;
    Iby_ATTR :	BYTE;
    Iby_BORDER :	BYTE;
    Xus_TN_SCREEN :	us_TN_SCREEN;

    func_block : TN_SC_LINE_Block;
	END_VAR
	func_block.Iin_X1 := Iin_X1;
	func_block.Iin_Y1 := Iin_Y1;
  func_block.Iin_X2 := Iin_X2;
	func_block.Iin_Y2 := Iin_Y2;
  func_block.Iby_ATTR := Iby_ATTR;
	func_block.Iby_BORDER := Iby_BORDER;
	func_block.Xus_TN_SCREEN := Xus_TN_SCREEN;

	func_block();
	Xus_TN_SCREEN  := func_block.Xus_TN_SCREEN;
END_PROGRAM

CONFIGURATION Config0
	RESOURCE Res0 ON PLC
		TASK task0(INTERVAL := T#20ms,PRIORITY := 0);
		PROGRAM instance0 WITH task0 : program0;
	END_RESOURCE
END_CONFIGURATION

(* ---- 690-YAHOO_WEATHER.ST ---- *)
FUNCTION_BLOCK YAHOO_WEATHER

  VAR_IN_OUT
    IP_C :	oscat_IP_C;
    S_BUF :	oscat_NETWORK_BUFFER;
    R_BUF :	oscat_NETWORK_BUFFER;
    YW :	oscat_YAHOO_WEATHER_DATA;
  END_VAR

  VAR_INPUT
    ACTIVATE :	BOOL;
    UNITS :	BOOL;
    LOCATION :	oscat_STRING20;
  END_VAR

  VAR_OUTPUT
    BUSY :	BOOL;
    DONE :	BOOL;
    ERROR_C :	DWORD;
    ERROR_T :	BYTE;
  END_VAR

  VAR
    CTRL :	oscat_XML_CONTROL;
    XML_READER :	XML_READER;
    URL_DATA :	oscat_url;
    DNS_CLIENT :	DNS_CLIENT;
    STRING_TO_URL :	STRING_TO_URL;
    HTTP_GET :	HTTP_GET;
    FLOAT_TO_REAL :	FLOAT_TO_REAL;
    CHK_REAL :	CHK_REAL;
    last_state :	BOOL;
    value_int :	INT;
    value_real :	REAL;
    v_real :	REAL;
    state :	INT;
  END_VAR

  CASE state OF

  00:
    IF ACTIVATE AND NOT last_state THEN
      state := 20;
    DONE := FALSE;
    BUSY := TRUE;
    ERROR_C := DWORD#0;
    ERROR_T := BYTE#0;
    END_IF;

  20:
    STRING_TO_URL.STR:='http://weather.yahooapis.com/forecastrss';
    STRING_TO_URL.DEFAULT_PROTOCOL:='';
    STRING_TO_URL.DEFAULT_PATH:='';
    STRING_TO_URL();
    URL_DATA:=STRING_TO_URL.STRING_TO_URL;

    URL_DATA.QUERY := CONCAT('w=',LOCATION);

    IF UNITS THEN
      URL_DATA.QUERY := CONCAT(URL_DATA.QUERY,'&u=f');
    ELSE
      URL_DATA.QUERY := CONCAT(URL_DATA.QUERY,'&u=c');
    END_IF;

    state := 40;

  40:
    IF DNS_CLIENT.DONE THEN
      state := 60;
    ELSIF (DNS_CLIENT.ERROR > DWORD#00) THEN
      ERROR_C := DNS_CLIENT.ERROR;
    ERROR_T := BYTE#01;
      state   := 100;
    END_IF;

  60:
    IF HTTP_GET.DONE THEN
      state := 80;
      CTRL.START_POS := HTTP_GET.BODY_START;
      CTRL.STOP_POS  := HTTP_GET.BODY_STOP;
      CTRL.COMMAND   := WORD#2#10000000_00011000;
    CTRL.WATCHDOG  := T#1ms;

    ELSIF (HTTP_GET.ERROR > DWORD#00) THEN
      ERROR_C := HTTP_GET.ERROR;
      ERROR_T := BYTE#02;
      state   := 100;
    END_IF;

  80:
    XML_READER.CTRL := CTRL;
    XML_READER.BUF  := R_BUF.BUFFER;
    XML_READER();
    CTRL         := XML_READER.CTRL;
    R_BUF.BUFFER := XML_READER.BUF;

    IF CTRL.TYP < 98 THEN
      value_int := 0;
    value_real := 0.0;
    IF LEN(CTRL.VALUE) <= 20 THEN
        FLOAT_TO_REAL(FLT:=CTRL.VALUE);
        v_real:=FLOAT_TO_REAL.FLOAT_TO_REAL;
      CHK_REAL(X:= v_real);
      IF CHK_REAL.CHK_REAL = BYTE#0 THEN
        value_real := v_real;
      value_int := REAL_TO_INT(value_real);
      END_IF;
    END_IF;

      IF CTRL.COUNT < UINT#52 THEN
        CASE UINT_TO_INT(CTRL.COUNT) OF
          027: YW.TimeToLive := value_int;
          030: YW.location_city := CTRL.VALUE;
          031: YW.location_region := CTRL.VALUE;
          032: YW.location_country := CTRL.VALUE;
          035: YW.unit_temperature := CTRL.VALUE;
          036: YW.unit_distance := CTRL.VALUE;
          037: YW.unit_pressure := CTRL.VALUE;
          038: YW.unit_speed := CTRL.VALUE;
          041: YW.wind_chill := value_int;
          042: YW.wind_direction := value_int;
          043: YW.wind_speed := value_real;
          046: YW.atmosphere_humidity := value_int;
          047: YW.atmosphere_visibility := value_real;
          048: YW.atmosphere_pressure := value_int;
          049: YW.atmosphere_rising := value_int;
        END_CASE;
      ELSE
        CASE UINT_TO_INT(CTRL.COUNT) OF
          052: YW.astronomy_sunrise := CTRL.VALUE;
          053: YW.astronomy_sunset := CTRL.VALUE;
          077: YW.geo_latitude := value_real;
          080: YW.geo_longitude := value_real;
          089: YW.cur_conditions_text := CTRL.VALUE;
      090: YW.cur_conditions_code := value_int;
        YW.cur_conditions_icon := value_int;
          091: YW.cur_conditions_temp := value_int;
          100: YW.forcast_today_low_temp := value_int;
          101: YW.forcast_today_high_temp := value_int;
          102: YW.forcast_today_text := CTRL.VALUE;
      103: YW.forcast_today_code := value_int;
        YW.forcast_today_icon := value_int;
          108: YW.forcast_tomorrow_low_temp := value_int;
          109: YW.forcast_tomorrow_high_temp := value_int;
          110: YW.forcast_tomorrow_text := CTRL.VALUE;
      111: YW.forcast_tomorrow_code := value_int;
        YW.forcast_tomorrow_icon := value_int;
        END_CASE;
      END_IF;
    ELSIF CTRL.TYP = 99 THEN
      DONE  := TRUE;
      state := 100;
    END_IF;

  100:
    IF (NOT HTTP_GET.DONE) THEN
      state := 0;
      BUSY  := FALSE;
      DONE := ERROR_T = BYTE#0;
    END_IF;

  END_CASE;

  DNS_CLIENT.IP_C     := IP_C;
  DNS_CLIENT.S_BUF    := S_BUF;
  DNS_CLIENT.R_BUF    := R_BUF;
  DNS_CLIENT.DOMAIN   := URL_DATA.DOMAIN;
  DNS_CLIENT.IP4_DNS  := DWORD#00;
  DNS_CLIENT.ACTIVATE := state=40;
  DNS_CLIENT();
  IP_C  := DNS_CLIENT.IP_C;
  S_BUF := DNS_CLIENT.S_BUF;
  R_BUF := DNS_CLIENT.R_BUF;

  HTTP_GET.IP_C        := IP_C;
  HTTP_GET.S_BUF       := S_BUF;
  HTTP_GET.R_BUF       := R_BUF;
  HTTP_GET.IP4         := DNS_CLIENT.IP4;
  HTTP_GET.GET         := state=60;
  HTTP_GET.MODE        := BYTE#2;
  HTTP_GET.UNLOCK_BUF  := state=100;
  HTTP_GET.URL_DATA    := URL_DATA;
  HTTP_GET();
  IP_C     := HTTP_GET.IP_C;
  S_BUF    := HTTP_GET.S_BUF;
  R_BUF    := HTTP_GET.R_BUF;
  URL_DATA := HTTP_GET.URL_DATA;

  last_state := ACTIVATE;

END_FUNCTION_BLOCK

(* ---- 691-ESR_MON_B8.ST ---- *)
TYPE
	oscat_esr_collect_data      : ARRAY [0..7]    OF BYTE;
END_TYPE
TYPE oscat_esr_data :
  STRUCT
	typ    : BYTE;
	adress : STRING;
	DS     : UDINT;
	TS     : TIME;
	data   : oscat_esr_collect_data;
  END_STRUCT;
END_TYPE

TYPE
  oscat_ESR_3                : ARRAY [0..3] OF oscat_esr_data;
  oscat_ESR_31               : ARRAY [0..31] OF oscat_esr_data;
END_TYPE

FUNCTION_BLOCK T_PLC_MS_block

	VAR_OUTPUT
		T_PLC_MS :	UDINT;
	END_VAR

	VAR_EXTERNAL
		PLC_TICKS_PER_SEC :	INT;
		PLC_SYS_TICK_CNT :	DINT;
	END_VAR

	VAR
		debug :	BOOL;(*Debug-Mode ON / OFF*)
		N :	INT;(*Debug-Faktor*)
		Offset :	UDINT;(*Debug-Offset*)
		temp :	DWORD := DWORD#1;(*Debug-Offset*)
		mode :	BOOL;(*modus*)
		faktor :	UDINT;(*Systemtakt-Faktor*)
		init :	BOOL;
		v_plc_ticks_per_sec :	UDINT;
		base :	UDINT := UDINT#1000;
	END_VAR

	IF init = FALSE THEN
		v_plc_ticks_per_sec := INT_TO_UDINT(PLC_TICKS_PER_SEC);
		IF v_plc_ticks_per_sec = UDINT#1024 THEN
			faktor := UDINT#1;
			mode := FALSE;
		ELSIF v_plc_ticks_per_sec > UDINT#0 THEN
			IF v_plc_ticks_per_sec <= base THEN
				faktor := base / v_plc_ticks_per_sec;
				mode := FALSE;
			ELSE
				faktor := v_plc_ticks_per_sec / base;
				mode := TRUE;
			END_IF;
		ELSE
			faktor := UDINT#1;
		END_IF;
		init := TRUE;
	END_IF;

	IF mode THEN
		T_PLC_MS := DINT_TO_UDINT(PLC_SYS_TICK_CNT) / faktor;
	ELSE
		T_PLC_MS := DINT_TO_UDINT(PLC_SYS_TICK_CNT) * faktor;
	END_IF;

	IF debug THEN
		T_PLC_MS := (DWORD_TO_UDINT(SHL(UDINT_TO_DWORD(T_PLC_MS),N) OR SHL(temp,N)) - UDINT#1) + Offset;
	END_IF;

END_FUNCTION_BLOCK

FUNCTION_BLOCK ESR_MON_B8

	VAR_INPUT
		S0 :	BOOL;
		A0 :	STRING;
		S1 :	BOOL;
		A1 :	STRING;
		S2 :	BOOL;
		A2 :	STRING;
		S3 :	BOOL;
		A3 :	STRING;
		S4 :	BOOL;
		A4 :	STRING;
		S5 :	BOOL;
		A5 :	STRING;
		S6 :	BOOL;
		A6 :	STRING;
		S7 :	BOOL;
		A7 :	STRING;
		DT_IN :	UDINT;
	END_VAR

	VAR_IN_OUT
		ESR_Out :	oscat_ESR_3;
	END_VAR

	VAR_OUTPUT
		ESR_FLAG :	BOOL;
	END_VAR

	VAR
		x0 :	BOOL;
		x1 :	BOOL;
		x2 :	BOOL;
		x3 :	BOOL;
		x4 :	BOOL;
		x5 :	BOOL;
		x6 :	BOOL;
		x7 :	BOOL;
		tx :	TIME;
		cnt :	INT;
		T_PLC_MS :	T_PLC_MS_block;
	END_VAR

	T_PLC_MS();
	tx:= UDINT_TO_TIME(T_PLC_MS.T_PLC_MS);

	ESR_Flag := FALSE;
	esr_out[3].typ := BYTE#0;
	esr_out[2].typ := BYTE#0;
	esr_out[1].typ := BYTE#0;
	esr_out[0].typ := BYTE#0;
	cnt := 0;

	IF s0 <> X0 THEN
		esr_out[cnt].typ := INT_TO_BYTE(10 + BOOL_TO_INT(s0));
		esr_out[cnt].adress := a0;
		esr_out[cnt].DS := DT_in;
		esr_out[cnt].TS := TX;
		X0 := S0;
		cnt := cnt + 1;
		esr_flag := TRUE;
	END_IF;
	IF s1 <> X1 THEN
		esr_out[cnt].typ := INT_TO_BYTE(10 + BOOL_TO_INT(s1));
		esr_out[cnt].adress := a1;
		esr_out[cnt].DS := DT_in;
		esr_out[cnt].TS := TX;
		X1 := S1;
		cnt := cnt + 1;
		esr_flag := TRUE;
	END_IF;
	IF s2 <> X2 THEN
		esr_out[cnt].typ := INT_TO_BYTE(10 + BOOL_TO_INT(s2));
		esr_out[cnt].adress := a2;
		esr_out[cnt].DS := DT_in;
		esr_out[cnt].TS := TX;
		X2 := S2;
		cnt := cnt + 1;
		esr_flag := TRUE;
	END_IF;
	IF s3 <> X3 THEN
		esr_out[cnt].typ := INT_TO_BYTE(10 + BOOL_TO_INT(s3));
		esr_out[cnt].adress := a3;
		esr_out[cnt].DS := DT_in;
		esr_out[cnt].TS := TX;
		X3 := S3;
		cnt := cnt + 1;
		esr_flag := TRUE;
	END_IF;
	IF s4 <> X4 AND cnt < 4 THEN
		esr_out[cnt].typ := INT_TO_BYTE(10 + BOOL_TO_INT(s4));
		esr_out[cnt].adress := a4;
		esr_out[cnt].DS := DT_in;
		esr_out[cnt].TS := TX;
		X4 := S4;
		cnt := cnt + 1;
		esr_flag := TRUE;
	END_IF;
	IF s5 <> X5  AND cnt < 4 THEN
		esr_out[cnt].typ := INT_TO_BYTE(10 + BOOL_TO_INT(s5));
		esr_out[cnt].adress := a5;
		esr_out[cnt].DS := DT_in;
		esr_out[cnt].TS := TX;
		X5 := S5;
		cnt := cnt + 1;
		esr_flag := TRUE;
	END_IF;
	IF s6 <> X6  AND cnt < 4 THEN
		esr_out[cnt].typ := INT_TO_BYTE(10 + BOOL_TO_INT(s6));
		esr_out[cnt].adress := a6;
		esr_out[cnt].DS := DT_in;
		esr_out[cnt].TS := TX;
		X6 := S6;
		cnt := cnt + 1;
		esr_flag := TRUE;
	END_IF;
	IF s7 <> X7  AND cnt < 4 THEN
		esr_out[cnt].typ := INT_TO_BYTE(10 + BOOL_TO_INT(s7));
		esr_out[cnt].adress := a7;
		esr_out[cnt].DS := DT_in;
		esr_out[cnt].TS := TX;
		X7 := S7;
		cnt := cnt + 1;
		esr_flag := TRUE;
	END_IF;

END_FUNCTION_BLOCK

PROGRAM program0

	VAR

		S0 :	BOOL;
		A0 :	STRING;
		S1 :	BOOL;
		A1 :	STRING;
		S2 :	BOOL;
		A2 :	STRING;
		S3 :	BOOL;
		A3 :	STRING;
		S4 :	BOOL;
		A4 :	STRING;
		S5 :	BOOL;
		A5 :	STRING;
		S6 :	BOOL;
		A6 :	STRING;
		S7 :	BOOL;
		A7 :	STRING;
		DT_IN   :	UDINT;

		ESR_Out :	oscat_ESR_3;

		ESR_FLAG :	BOOL;

		func_block : ESR_MON_B8;
  	END_VAR
	func_block.S0 := S0;
	func_block.A0 := A0;
	func_block.S1 := S1;
	func_block.A1 := A1;
	func_block.S2 := S2;
	func_block.A2 := A2;
	func_block.S3 := S3;
	func_block.A3 := A3;
	func_block.S4 := S4;
	func_block.A4 := A4;
	func_block.S5 := S5;
	func_block.A5 := A5;
	func_block.S6 := S6;
	func_block.A6 := A6;
	func_block.S7 := S7;
	func_block.A7 := A7;
	func_block.DT_IN := DT_IN;
	func_block.ESR_Out := ESR_Out;
	func_block();
	ESR_Out := func_block.ESR_Out;
	ESR_FLAG := func_block.ESR_FLAG;

END_PROGRAM

CONFIGURATION Config0

	VAR_GLOBAL
		PLC_TICKS_PER_SEC :	INT;
		PLC_SYS_TICK_CNT :	DINT;
	END_VAR

  	RESOURCE Res0 ON PLC
    	TASK task0(INTERVAL := T#20ms,PRIORITY := 0);
    	PROGRAM instance0 WITH task0 : program0;
  	END_RESOURCE

END_CONFIGURATION

(* ---- 692-DT_TO_STRF.ST ---- *)
FUNCTION DT_TO_DATE2:UDINT

	VAR_INPUT
		IN :	UDINT;
	END_VAR

	DT_TO_DATE2 := (IN / UDINT#86400) * UDINT#86400;
END_FUNCTION

FUNCTION DT_TO_TOD2:UDINT
	VAR_INPUT
		IN :	UDINT;
	END_VAR

	DT_TO_TOD2 := (IN MOD UDINT#86400) * UDINT#1000;
END_FUNCTION

FUNCTION _BYTE_TO_INT:INT
	VAR_INPUT
		IN :	BYTE;
	END_VAR

	_BYTE_TO_INT := USINT_TO_INT(BYTE_TO_USINT(IN));
END_FUNCTION

FUNCTION_BLOCK DT_TO_STRF_Block

	VAR_INPUT
		DTI :	UDINT;
		MS :	INT;
		FMT :	STRING;
		LANG :	INT;
	END_VAR

	VAR_OUTPUT
		DT_TO_STRF :	STRING;
	END_VAR

	VAR
		FILL :	STRING;
		BLANK :	STRING;
		ly :	INT;
		dx :	UDINT;
		fs :	STRING;
		fs_tmp :	STRING;
		td :	UDINT;
		tmp :	INT;
		pos :	INT;
		f :	INT;
		CODEE :	CODE;
		MONTH_TO_STRING :	MONTH_TO_STRING;
		WEEKDAY_TO_STRING :	WEEKDAY_TO_STRING;
	END_VAR

	IF LANG < 1 THEN ly := 1; ELSE ly := MIN(2, LANG); END_IF;

	dx := DT_TO_DATE2(DTI);
	td := DT_TO_TOD2(DTI);

	DT_TO_STRF := FMT;
	pos := FIND(DT_TO_STRF, '#');
	WHILE pos > 0 DO
		CODEE(STR:=DT_TO_STRF,POS:=pos + 1);
		f := _BYTE_TO_INT(CODEE.CODEE);
		(* generate the return string according to the format character *)
		fs := '';
		CASE f OF
			0: RETURN; (* illegal character index *)

			65 : (* letter A retunrs the year in 4 digits *)
				fs := INT_TO_STRING(YEAR_OF_DATE(dx),'%d');
			66 : (* letter B returns the year in exactly 2 digits *)
				fs := RIGHT(INT_TO_STRING(YEAR_OF_DATE(dx),'%02d'),2);
			67 : (* letter C returns the month with 1 or 2 digits *)
				fs := INT_TO_STRING(MONTH_OF_DATE(dx),'%d');
			68 : (* letter D returns the month with exactly 2 digits *)
				fs := INT_TO_STRING(MONTH_OF_DATE(dx),'%02d');
			69 : (* letter E returns the month with 3 characters *)
				MONTH_TO_STRING(MTH:=MONTH_OF_DATE(dx),LANG:=ly,LX:=3);
				fs:=MONTH_TO_STRING.MONTH_TO_STRING;
			70 : (* letter F returns the month with all characters *)
				MONTH_TO_STRING(MTH:=MONTH_OF_DATE(dx),LANG:=ly,LX:=0);
				fs:=MONTH_TO_STRING.MONTH_TO_STRING;
			71 : (* letter G returns the day with up to 2 digits *)
				fs := INT_TO_STRING(DAY_OF_MONTH(dx),'%d');
			72 : (* letter H returns the day of the month with exactly 2 digits *)
				fs := INT_TO_STRING(DAY_OF_MONTH(dx),'%d');
				IF LEN(fs) < 2 THEN fs_tmp:=fs; fs := CONCAT(FILL, fs_tmp); END_IF;
			73 : (* letter I returns the weekday as the number 1..7 1 = monday *)
				fs := INT_TO_STRING(DAY_OF_WEEK(dx),'%d');
			74 : (* letter J returns the weekday in 2 character writing *)
				WEEKDAY_TO_STRING(WDAY:=DAY_OF_WEEK(dx),LANG:=ly,LX:=2);
				fs := WEEKDAY_TO_STRING.WEEKDAY_TO_STRING;
			75 : (* letter K returns the weekday with all characters *)
				WEEKDAY_TO_STRING(WDAY:=DAY_OF_WEEK(dx),LANG:=ly,LX:=0);
				fs := WEEKDAY_TO_STRING.WEEKDAY_TO_STRING;
			76 : (* letter L returns AM or PM for the given DateTime *)
				IF td >= UDINT#43200000 THEN fs := 'PM'; ELSE fs := 'AM'; END_IF;
			77 : (* letter M returns the hour in 1 or 2 digit form 0..24h *)
				fs := INT_TO_STRING(HOUR(td),'%d');
			78 : (* letter N returns the hour in exactly 2 digit form 0..24h *)
				fs := INT_TO_STRING(HOUR(td),'%d');
				IF LEN(fs) < 2 THEN fs_tmp:=fs; fs := CONCAT(FILL, fs_tmp); END_IF;
			79 : (* letter O returns the hour in 1 or 2 digit form 0..12h *)
				tmp := HOUR(td) MOD 12;
				IF tmp = 0 THEN tmp := 12; END_IF;
				fs := INT_TO_STRING(tmp,'%d');
			80 : (* letter P returns the hour in exactly 2 digit form 0..12h *)
				tmp := HOUR(td) MOD 12;
				IF tmp = 0 THEN tmp := 12; END_IF;
				fs := INT_TO_STRING(tmp,'%d');
				IF LEN(fs) < 2 THEN fs_tmp:=fs; fs := CONCAT(FILL, fs_tmp); END_IF;
			81 : (* letter Q returns the minute of the hour in 1 or two digit form *)
				fs := INT_TO_STRING(MINUTE(td),'%d');
			82 : (* letter R returns the minute of the hour in exactly two digit form *)
				fs := INT_TO_STRING(MINUTE(td),'%d');
				IF LEN(fs) < 2 THEN fs_tmp:=fs; fs := CONCAT(FILL, fs_tmp); END_IF;
			83 : (* letter S returns the second of the minute in 1 or two digit form *)
				fs := INT_TO_STRING(REAL_TO_INT(SECOND(td)),'%d');
			84 : (* letter T returns the second of the minute in exactly two digit form *)
				fs := INT_TO_STRING(REAL_TO_INT(SECOND(td)),'%d');
				IF LEN(fs) < 2 THEN fs_tmp:=fs; fs := CONCAT(FILL, fs_tmp); END_IF;
			85 : (* letter U returns the milliseconds in 1 to 3 digits *)
				fs := INT_TO_STRING(MS,'%d');
			86 : (* letter V returns the milliseconds in exactly 3 digit form *)
				fs := INT_TO_STRING(MS,'%03d');
			87 : (* letter W returns the day of the month with exactly 2 digits first digit is filled with blank if necessary *)
				fs := INT_TO_STRING(DAY_OF_MONTH(dx),'%d');
				IF LEN(fs) < 2 THEN fs_tmp:=fs; fs := CONCAT(BLANK, fs_tmp); END_IF;
			88 : (* letter X returns the month with exactly 2 digits first digit is filled with blank if necessary *)
				fs := INT_TO_STRING(MONTH_OF_DATE(dx),'%d');
				IF LEN(fs) < 2 THEN fs_tmp:=fs; fs := CONCAT(BLANK, fs_tmp); END_IF;
		END_CASE;
		DT_TO_STRF := REPLACE(DT_TO_STRF, fs, 2, pos);
		pos := FIND(DT_TO_STRF, '#');
	END_WHILE;

END_FUNCTION_BLOCK

PROGRAM program0
  VAR
	DTI  :	UDINT;
	MS   :	INT;
	FMT  :	STRING;
	LANG :	INT;

	DT_TO_STRF :	STRING;

	func_block : DT_TO_STRF_Block;
  END_VAR
	func_block.DTI  :=DTI ;
	func_block.MS   :=MS  ;
	func_block.FMT  :=FMT ;
	func_block.LANG :=LANG;
	func_block();
	DT_TO_STRF := func_block.DT_TO_STRF;
END_PROGRAM

CONFIGURATION Config0
  RESOURCE Res0 ON PLC
    TASK task0(INTERVAL := T#20ms,PRIORITY := 0);
    PROGRAM instance0 WITH task0 : program0;
  END_RESOURCE
END_CONFIGURATION

(* ---- 693-ACTUATOR_2P.ST ---- *)
FUNCTION UDINT_TO_TIME2:TIME

	VAR_INPUT
		IN :	UDINT;
	END_VAR

	UDINT_TO_TIME2 := DINT_TO_TIME(UDINT_TO_DINT(IN));

END_FUNCTION

FUNCTION_BLOCK T_PLC_MS_block
	VAR_OUTPUT
		T_PLC_MS :	UDINT;
	END_VAR

	VAR_EXTERNAL
		PLC_TICKS_PER_SEC :	INT;
		PLC_SYS_TICK_CNT :	DINT;
	END_VAR

	VAR
		debug :	BOOL;(*Debug-Mode ON / OFF*)
		N :	INT;(*Debug-Faktor*)
		Offset :	UDINT;(*Debug-Offset*)
		temp :	DWORD := DWORD#1;(*Debug-Offset*)
		mode :	BOOL;(*modus*)
		faktor :	UDINT;(*Systemtakt-Faktor*)
		init :	BOOL;
		v_plc_ticks_per_sec :	UDINT;
		base :	UDINT := UDINT#1000;
	END_VAR

	IF init = FALSE THEN
		v_plc_ticks_per_sec := INT_TO_UDINT(PLC_TICKS_PER_SEC);
		IF v_plc_ticks_per_sec = UDINT#1024 THEN
			faktor := UDINT#1;
			mode := FALSE;
		ELSIF v_plc_ticks_per_sec > UDINT#0 THEN
			IF v_plc_ticks_per_sec <= base THEN
				faktor := base / v_plc_ticks_per_sec;
				mode := FALSE;
			ELSE
				faktor := v_plc_ticks_per_sec / base;
				mode := TRUE;
			END_IF;
		ELSE
			faktor := UDINT#1;
		END_IF;
		init := TRUE;
	END_IF;

	IF mode THEN
		T_PLC_MS := DINT_TO_UDINT(PLC_SYS_TICK_CNT) / faktor;
	ELSE
		T_PLC_MS := DINT_TO_UDINT(PLC_SYS_TICK_CNT) * faktor;
	END_IF;

	IF debug THEN
		T_PLC_MS := (DWORD_TO_UDINT(SHL(UDINT_TO_DWORD(T_PLC_MS),N) OR SHL(temp,N)) - UDINT#1) + Offset;
	END_IF;

END_FUNCTION_BLOCK

FUNCTION TIME_TO_UDINT2:UDINT
	VAR_INPUT
		X :	TIME;
	END_VAR

	TIME_TO_UDINT2 := DINT_TO_UDINT(TIME_TO_DINT(X));
END_FUNCTION

FUNCTION FRMP_B:BYTE
	VAR_INPUT
		START :	BYTE;
		DIR :	BOOL;
		TD :	TIME;
		TR :	TIME;
	END_VAR

	IF TD < TR THEN
		FRMP_B := MIN(UDINT_TO_BYTE(DWORD_TO_UDINT(SHL(TIME_TO_DWORD(TD), 8)) / TIME_TO_UDINT2(TR)), SEL(DIR, START, USINT_TO_BYTE(USINT#255 - BYTE_TO_USINT(START))));
		IF DIR THEN
			FRMP_B := USINT_TO_BYTE(BYTE_TO_USINT(START) + BYTE_TO_USINT(FRMP_B));
		ELSE
			FRMP_B := USINT_TO_BYTE(BYTE_TO_USINT(START) - BYTE_TO_USINT(FRMP_B));
		END_IF;
	ELSE
		FRMP_B := SEL(DIR, BYTE#0, BYTE#255);
	END_IF;
END_FUNCTION

FUNCTION_BLOCK _RMP_B
	VAR_INPUT
		DIR :	BOOL;
		E :	BOOL := TRUE;
		TR :	TIME;
	END_VAR

	VAR_IN_OUT
		RMP :	BYTE;
	END_VAR

	VAR
		T_PLC_MS :	T_PLC_MS_block;
		tx :	TIME;
		tl :	TIME;
		tn :	TIME;
		init :	BOOL;
		last_dir :	BOOL;
		start :	BYTE;
	END_VAR

	T_PLC_MS();
	tx := UDINT_TO_TIME(T_PLC_MS.T_PLC_MS);

	IF E AND init AND (dir = last_dir) AND (RMP <> SEL(DIR, BYTE#0, BYTE#255)) AND TR = tn THEN
		RMP := FRMP_B(start, DIR, tx - tl, TR);
	ELSE
		init := TRUE;
		tl := tx;
		tn := tr;
		start := RMP;
	END_IF;
	last_dir := dir;
END_FUNCTION_BLOCK

FUNCTION_BLOCK AUTORUN_Block

	VAR_INPUT
		IN :	BOOL;
		TEST :	BOOL;
		ARE :	BOOL := TRUE;
		TRUN :	TIME;
		TOFF :	TIME;
	END_VAR

	VAR_OUTPUT
		OUT :	BOOL;
		ARO :	BOOL;
	END_VAR

	VAR_IN_OUT
		ARX :	BOOL;
	END_VAR

	VAR
		timer :	_RMP_B;
		val :	BYTE;
	END_VAR

	IF TOFF > T#0s THEN
		timer(DIR:= OUT, TR := SEL(OUT, TOFF, TRUN), RMP := val);
		val := timer.RMP;
	ELSE
		val := BYTE#255;
	END_IF;

	IF (NOT ARX AND ARE AND val = BYTE#0) OR TEST THEN
		val := BYTE#0;
		ARO := TRUE;
		ARX := TRUE;
	ELSIF val = BYTE#255 AND ARO THEN
		ARO := FALSE;
		ARX := FALSE;
	END_IF;

	out := IN OR ARO;

END_FUNCTION_BLOCK

FUNCTION_BLOCK GEN_PULSE_Block

	VAR_INPUT
		ENQ :	BOOL := TRUE;
		PTH :	TIME;
		PTL :	TIME;
	END_VAR

	VAR_OUTPUT
		Q :	BOOL;
	END_VAR

	VAR
		T_PLC_MS :	T_PLC_MS_block;
		tx :	TIME;
		tn :	TIME;
		init :	BOOL;
	END_VAR

	IF enq THEN
		T_PLC_MS();
		tx:= UDINT_TO_TIME(T_PLC_MS.T_PLC_MS);
		IF NOT init THEN init := TRUE; tn := tx; END_IF;
		IF tx - tn >= SEL(Q, PTL, PTH) THEN
			tn := tn + SEL(Q, PTL, PTH);
			Q := NOT Q;
		END_IF;
	ELSE
		Q := FALSE;
		init := FALSE;
	END_IF;

END_FUNCTION_BLOCK

FUNCTION_BLOCK ACTUATOR_2P_Block

	VAR_INPUT
		IN :	BYTE;
		TEST :	BOOL;
		ARE :	BOOL := TRUE;
		CYCLE_TIME :	TIME;
		SENS :	BYTE;
		SELF_ACT_TIME :	TIME;
		SELF_ACT_PULSE :	TIME;
		SELF_ACT_CYCLES :	INT := 1;
	END_VAR

	VAR_OUTPUT
		OUT :	BOOL;
		ARO :	BOOL;
	END_VAR

	VAR_IN_OUT
		ARX :	BOOL;
	END_VAR

	VAR
		timer :	AUTORUN_Block;
		pwgen :	GEN_PULSE_Block;
	END_VAR

	timer(trun := MUL_T_AI(SELF_ACT_PULSE,2 * SELF_ACT_CYCLES), toff := SELF_ACT_TIME, Test := TEST, ARE := ARE, arx := ARX);
	ARX := timer.ARX;
	ARO := timer.ARO;

	IF aro THEN
		pwgen(PTL := SELF_ACT_PULSE, PTH := SELF_ACT_PULSE);
		out := pwgen.Q;
	ELSIF in < sens THEN
		out := FALSE;
	ELSIF BYTE_TO_USINT(in) > USINT#255 - BYTE_TO_USINT(sens) THEN
		out := TRUE;
	ELSE
		pwgen.PTH := (CYCLE_TIME * BYTE_TO_TIME2(BAND_B(IN,SENS))  ) / BYTE_TO_TIME2(BYTE#255);
		pwgen.PTL := CYCLE_TIME - pwgen.PTH;
		pwgen();
		out := pwgen.Q;
	END_IF;

END_FUNCTION_BLOCK

PROGRAM program0
	VAR
		IN :	BYTE;
		TEST :	BOOL;
		ARE :	BOOL := TRUE;
		CYCLE_TIME :	TIME;
		SENS :	BYTE;
		SELF_ACT_TIME :	TIME;
		SELF_ACT_PULSE :	TIME;
		SELF_ACT_CYCLES :	INT := 1;
		OUT :	BOOL;
		ARO :	BOOL;
		func_block : ACTUATOR_2P_Block;
	END_VAR
	func_block.IN := IN;
	func_block.TEST := TEST;
	func_block.ARE := ARE ;
	func_block.CYCLE_TIME := CYCLE_TIME;
	func_block.SENS := SENS;
	func_block.SELF_ACT_TIME := SELF_ACT_TIME ;
	func_block.SELF_ACT_PULSE := SELF_ACT_PULSE;
	func_block.SELF_ACT_CYCLES := SELF_ACT_CYCLES;
	func_block();
	OUT  := func_block.OUT;
	ARO  := func_block.ARO;
END_PROGRAM

CONFIGURATION Config0
	VAR_GLOBAL
		PLC_TICKS_PER_SEC :	INT;
		PLC_SYS_TICK_CNT :	DINT;
	END_VAR
  	RESOURCE Res0 ON PLC
    	TASK task0(INTERVAL := T#20ms,PRIORITY := 0);
    	PROGRAM instance0 WITH task0 : program0;
  	END_RESOURCE
END_CONFIGURATION

(* ---- 694-FT_PROFILE.ST ---- *)
FUNCTION_BLOCK T_PLC_MS_block
	VAR_OUTPUT
		T_PLC_MS :	UDINT;
	END_VAR

	VAR_EXTERNAL
		PLC_TICKS_PER_SEC :	INT;
		PLC_SYS_TICK_CNT :	DINT;
	END_VAR

	VAR
		debug :	BOOL;(*Debug-Mode ON / OFF*)
		N :	INT;(*Debug-Faktor*)
		Offset :	UDINT;(*Debug-Offset*)
		temp :	DWORD := DWORD#1;(*Debug-Offset*)
		mode :	BOOL;(*modus*)
		faktor :	UDINT;(*Systemtakt-Faktor*)
		init :	BOOL;
		v_plc_ticks_per_sec :	UDINT;
		base :	UDINT := UDINT#1000;
	END_VAR

	IF init = FALSE THEN
		v_plc_ticks_per_sec := INT_TO_UDINT(PLC_TICKS_PER_SEC);
		IF v_plc_ticks_per_sec = UDINT#1024 THEN
			faktor := UDINT#1;
			mode := FALSE;
		ELSIF v_plc_ticks_per_sec > UDINT#0 THEN
			IF v_plc_ticks_per_sec <= base THEN
				faktor := base / v_plc_ticks_per_sec;
				mode := FALSE;
			ELSE
				faktor := v_plc_ticks_per_sec / base;
				mode := TRUE;
			END_IF;
		ELSE
			faktor := UDINT#1;
		END_IF;
		init := TRUE;
	END_IF;

	IF mode THEN
		T_PLC_MS := DINT_TO_UDINT(PLC_SYS_TICK_CNT) / faktor;
	ELSE
		T_PLC_MS := DINT_TO_UDINT(PLC_SYS_TICK_CNT) * faktor;
	END_IF;

	IF debug THEN
		T_PLC_MS := (DWORD_TO_UDINT(SHL(UDINT_TO_DWORD(T_PLC_MS),N) OR SHL(temp,N)) - UDINT#1) + Offset;
	END_IF;
END_FUNCTION_BLOCK

FUNCTION_BLOCK FT_PROFILE

	VAR_INPUT
		K :	REAL := 1.0;
		O :	REAL := 0.0;
		M :	REAL := 1.0;
		E :	BOOL;
		VALUE_0 :	REAL;
		TIME_1 :	TIME;
		VALUE_1 :	REAL;
		TIME_2 :	TIME;
		VALUE_2 :	REAL;
		TIME_3 :	TIME;
		VALUE_3 :	REAL;
		TIME_10 :	TIME;
		VALUE_10 :	REAL;
		TIME_11 :	TIME;
		VALUE_11 :	REAL;
		TIME_12 :	TIME;
		VALUE_12 :	REAL;
		TIME_13 :	TIME;
		VALUE_13 :	REAL;
	END_VAR

	VAR_OUTPUT
		Y :	REAL;
		RUN :	BOOL;
		ET :	TIME;
	END_VAR

	VAR
		tx :	TIME;
		edge :	BOOL;
		state :	INT;
		ta :	TIME;
		tb :	TIME;
		t0 :	TIME;
		temp :	REAL;
		va :	REAL;
		vb :	REAL;
		T_PLC_MS :	T_PLC_MS_block;
	END_VAR

	T_PLC_MS();
	tx:= UDINT_TO_TIME(T_PLC_MS.T_PLC_MS);

	(* determine start condition *)
	IF E AND NOT edge THEN
		RUN := TRUE;
		ET := t#0s;
		t0 := tx;
		ta := tx;
		tb := multime(time_1, M);
		va := value_0;
		vb := value_1;
		temp := value_0;
		state := 1;
	END_IF;
	edge := E;

	(* generate startup profile *)
	IF run THEN
		CASE state OF
			1:	IF tx - ta >= tb THEN
					ta := ta + tb;
					tb := multime(time_2 - time_1, M);
					va := value_1;
					vb := value_2;
					temp := value_1;
					state := 2;
				ELSE
					temp := ((vb - va) * TIME_TO_REAL(tx - ta) / TIME_TO_REAL(tb) + va);
				END_IF;
			2:	IF tx - ta >= tb THEN
					ta := ta + tb;
					tb := multime(time_3 - time_2, M);
					va := value_2;
					vb := value_3;
					temp := value_2;
					state := 3;
				ELSE
					temp := ((vb - va) * TIME_TO_REAL(tx - ta) / TIME_TO_REAL(tb) + va);
				END_IF;
			3:	IF tx - ta >= tb THEN
					ta := ta + tb;
					tb := multime(time_10 - time_3, M);
					va := value_3;
					vb := value_10;
					temp := value_3;
					state := 4;
				ELSE
					temp := ((vb - va) * TIME_TO_REAL(tx - ta) / TIME_TO_REAL(tb) + va);
				END_IF;
			4 :	IF tx - ta >= tb THEN
					ta := ta + tb;
					tb := multime(time_11 - time_10, M);
					va := value_10;
					vb := value_11;
					temp := value_10;
					IF E THEN state := 5; ELSE state := 6; END_IF;
				ELSE
					temp := ((vb - va) * TIME_TO_REAL(tx - ta) / TIME_TO_REAL(tb) + va);
				END_IF;
			5:	(* extend the signal while E is true *)
				IF E THEN
					ta := tx;
				ELSE
					state := 6;
				END_IF;
			6:	IF tx - ta >= tb THEN
					ta := ta + tb;
					tb := multime(time_12 - time_11, M);
					va := value_11;
					vb := value_12;
					temp := value_11;
					state := 7;
				ELSE
					temp := ((vb - va) * TIME_TO_REAL(tx - ta) / TIME_TO_REAL(tb) + va);
				END_IF;
			7:	IF tx - ta >= tb THEN
					ta := ta + tb;
					tb := multime(time_13 - time_12, M);
					va := value_12;
					vb := value_13;
					temp := value_12;
					state := 8;
				ELSE
					temp := ((vb - va) * TIME_TO_REAL(tx - ta) / TIME_TO_REAL(tb) + va);
				END_IF;
			8:	IF tx - ta >= tb THEN
					temp := value_13;
					run := FALSE;
				ELSE
					temp := ((vb - va) * TIME_TO_REAL(tx - ta) / TIME_TO_REAL(tb) + va);
				END_IF;
		END_CASE;
		Y := temp * K + O;
		ET := tx - t0;
	END_IF;

END_FUNCTION_BLOCK

PROGRAM program0
	VAR
		K :	REAL := 1.0;
		O :	REAL := 0.0;
		M :	REAL := 1.0;
		E :	BOOL;
		VALUE_0 :	REAL;
		TIME_1 :	TIME;
		VALUE_1 :	REAL;
		TIME_2 :	TIME;
		VALUE_2 :	REAL;
		TIME_3 :	TIME;
		VALUE_3 :	REAL;
		TIME_10 :	TIME;
		VALUE_10 :	REAL;
		TIME_11 :	TIME;
		VALUE_11 :	REAL;
		TIME_12 :	TIME;
		VALUE_12 :	REAL;
		TIME_13 :	TIME;
		VALUE_13 :	REAL;

		Y :	REAL;
		RUN :	BOOL;
		ET :	TIME;

		func_block : FT_PROFILE;
	END_VAR
	func_block.K  := K ;
	func_block.O  := O ;
	func_block.M  := M ;
	func_block.E  := E ;
	func_block.VALUE_0  := VALUE_0 ;
	func_block.TIME_1  := TIME_1 ;
	func_block.VALUE_1  := VALUE_1 ;
	func_block.TIME_2  := TIME_2 ;
	func_block.VALUE_2  := VALUE_2 ;
	func_block.TIME_3  := TIME_3 ;
	func_block.VALUE_3  := VALUE_3 ;
	func_block.TIME_10  := TIME_10 ;
	func_block.VALUE_10  := VALUE_10 ;
	func_block.TIME_11  := TIME_11 ;
	func_block.VALUE_11  := VALUE_11 ;
	func_block.TIME_12  := TIME_12 ;
	func_block.VALUE_12  := VALUE_12 ;
	func_block.TIME_13  := TIME_13 ;
	func_block.VALUE_13  := VALUE_13 ;
	func_block();
	Y := func_block.Y;
	RUN := func_block.RUN;
	ET := func_block.ET;
END_PROGRAM

CONFIGURATION Config0

	VAR_GLOBAL
		PLC_TICKS_PER_SEC :	INT;
		PLC_SYS_TICK_CNT :	DINT;
	END_VAR

	RESOURCE Res0 ON PLC
		TASK task0(INTERVAL := T#20ms,PRIORITY := 0);
		PROGRAM instance0 WITH task0 : program0;
	END_RESOURCE

END_CONFIGURATION

(* ---- 695-GEN_RDT.ST ---- *)
FUNCTION _REAL_TO_UDINT:UDINT
  VAR_INPUT
    X :	REAL;
  END_VAR

  IF REAL_TO_UDINT(0.5) = UDINT#1 THEN
    _REAL_TO_UDINT := REAL_TO_UDINT(x);
  ELSIF X > 0.0 THEN
    _REAL_TO_UDINT := REAL_TO_UDINT(x+0.5);
  ELSIF X < 0.0 THEN
    _REAL_TO_UDINT := REAL_TO_UDINT(x-0.5);
  ELSE
    _REAL_TO_UDINT := UDINT#0;
  END_IF;
END_FUNCTION

FUNCTION REAL_TO_TIME2:TIME
	VAR_INPUT
		IN :	REAL;
	END_VAR

	REAL_TO_TIME2 := DINT_TO_TIME(UDINT_TO_DINT(_REAL_TO_UDINT(IN)));
END_FUNCTION

FUNCTION TIME_TO_REAL1:REAL

VAR_INPUT
	X :	TIME;
END_VAR

TIME_TO_REAL1 := UDINT_TO_REAL(DINT_TO_UDINT(TIME_TO_DINT(X)));
END_FUNCTION

FUNCTION D_TRUNC : DINT
  VAR_INPUT
    x : REAL;
  END_VAR

  D_TRUNC := REAL_TO_DINT(X);
  IF X > 0.0 THEN
  	IF DINT_TO_REAL(D_TRUNC) > X THEN D_TRUNC := D_TRUNC - DINT#1; END_IF;
  ELSE
  	IF DINT_TO_REAL(D_TRUNC) < X THEN D_TRUNC := D_TRUNC + DINT#1; END_IF;
  END_IF;
END_FUNCTION

FUNCTION BIT_COUNT:INT

	VAR_INPUT
		IN :	DWORD;
	END_VAR

	VAR
		in_temp :	DWORD;
	END_VAR

	in_temp := IN;
	WHILE in_temp > DWORD#0 DO
		IF (in_temp AND DWORD#16#00000001) > DWORD#0 THEN Bit_Count := Bit_Count +1; END_IF;
		in_temp := SHR(in_temp,1);
	END_WHILE;

END_FUNCTION

FUNCTION FRACT:REAL
	VAR_INPUT
		X :	REAL;
	END_VAR

	IF ABS(x) < 2.0E9 THEN
		FRACT := x - DINT_TO_REAL(D_TRUNC(x));
	ELSE
		FRACT := 0.0;
	END_IF;

END_FUNCTION

FUNCTION_BLOCK T_PLC_MS_block
	VAR_OUTPUT
		T_PLC_MS :	UDINT;
	END_VAR

	VAR_EXTERNAL
		PLC_TICKS_PER_SEC :	INT;
		PLC_SYS_TICK_CNT :	DINT;
	END_VAR

	VAR
		debug :	BOOL;(*Debug-Mode ON / OFF*)
		N :	INT;(*Debug-Faktor*)
		Offset :	UDINT;(*Debug-Offset*)
		temp :	DWORD := DWORD#1;(*Debug-Offset*)
		mode :	BOOL;(*modus*)
		faktor :	UDINT;(*Systemtakt-Faktor*)
		init :	BOOL;
		v_plc_ticks_per_sec :	UDINT;
		base :	UDINT := UDINT#1000;
	END_VAR

	IF init = FALSE THEN
		v_plc_ticks_per_sec := INT_TO_UDINT(PLC_TICKS_PER_SEC);
		IF v_plc_ticks_per_sec = UDINT#1024 THEN
			faktor := UDINT#1;
			mode := FALSE;
		ELSIF v_plc_ticks_per_sec > UDINT#0 THEN
			IF v_plc_ticks_per_sec <= base THEN
				faktor := base / v_plc_ticks_per_sec;
				mode := FALSE;
			ELSE
				faktor := v_plc_ticks_per_sec / base;
				mode := TRUE;
			END_IF;
		ELSE
			faktor := UDINT#1;
		END_IF;
		init := TRUE;
	END_IF;

	IF mode THEN
		T_PLC_MS := DINT_TO_UDINT(PLC_SYS_TICK_CNT) / faktor;
	ELSE
		T_PLC_MS := DINT_TO_UDINT(PLC_SYS_TICK_CNT) * faktor;
	END_IF;

	IF debug THEN
		T_PLC_MS := (DWORD_TO_UDINT(SHL(UDINT_TO_DWORD(T_PLC_MS),N) OR SHL(temp,N)) - UDINT#1) + Offset;
	END_IF;

END_FUNCTION_BLOCK

FUNCTION BIT_LOAD_DW:DWORD

	VAR_INPUT
		IN :	DWORD;
		VAL :	BOOL;
		POS :	INT;
	END_VAR

	IF val THEN
		BIT_LOAD_DW := in OR SHL(DWORD#1,pos);
	ELSE
		BIT_LOAD_DW := in AND (NOT SHL(DWORD#1,pos));
	END_IF;

END_FUNCTION

FUNCTION BIT_OF_DWORD : BOOL
  VAR_INPUT
    IN : DWORD;
    N : INT;
  END_VAR

  BIT_OF_DWORD := (SHR(in,N) AND 16#00000001) > 0;
  (* from OSCAT library; www.oscat.de  *)
END_FUNCTION

FUNCTION _INT_TO_UDINT:UDINT
	VAR_INPUT
		IN :	INT;
	END_VAR

	_INT_TO_UDINT := DINT_TO_UDINT(INT_TO_DINT(IN));
END_FUNCTION

FUNCTION _DWORD_TO_REAL:REAL
	VAR_INPUT
		IN :	DWORD;
	END_VAR

	_DWORD_TO_REAL := UDINT_TO_REAL(DWORD_TO_UDINT(IN));

END_FUNCTION

FUNCTION_BLOCK RDM_block
	VAR_INPUT
		LAST :	REAL;
	END_VAR
	VAR_OUTPUT
		RDM :	REAL;
	END_VAR
	VAR
		T_PLC_MS :	T_PLC_MS_block;
		tn :	DWORD;
		tc :	INT;
	END_VAR
	T_PLC_MS();
	tn := UDINT_TO_DWORD(T_PLC_MS.T_PLC_MS);
	tc := Bit_Count(tn);

	tn:=BIT_LOAD_DW(tn,BIT_OF_DWORD(tn,2),31); (* tn.31 := tn.2; *)
	tn:=BIT_LOAD_DW(tn,BIT_OF_DWORD(tn,5),30); (* tn.30 := tn.5; *)
	tn:=BIT_LOAD_DW(tn,BIT_OF_DWORD(tn,4),29); (* tn.29 := tn.4; *)
	tn:=BIT_LOAD_DW(tn,BIT_OF_DWORD(tn,1),28); (* tn.28 := tn.1; *)
	tn:=BIT_LOAD_DW(tn,BIT_OF_DWORD(tn,0),27); (* tn.27 := tn.0; *)
	tn:=BIT_LOAD_DW(tn,BIT_OF_DWORD(tn,7),26); (* tn.26 := tn.7; *)
	tn:=BIT_LOAD_DW(tn,BIT_OF_DWORD(tn,6),25); (* tn.25 := tn.6; *)
	tn:=BIT_LOAD_DW(tn,BIT_OF_DWORD(tn,3),24); (* tn.24 := tn.3; *)

	tn := ROL(tn,Bit_Count(tn)) OR DWORD#16#80000001;
	tn := UDINT_TO_DWORD(DWORD_TO_UDINT(tn) MOD UDINT#71474513 + _INT_TO_UDINT(tc) + UDINT#77);
	RDM := fract(_DWORD_TO_REAL(tn) / 10000000.0 * (2.71828182845904523536028747135266249 - LIMIT_REAL(0.0,last,1.0)));
END_FUNCTION_BLOCK

FUNCTION_BLOCK GEN_RDT_Block

	VAR_INPUT
		ENABLE :	BOOL := TRUE;
		MIN_TIME_MS :	TIME := t#1s;
		MAX_TIME_MS :	TIME := t#1.2s;
		TP_Q :	TIME := t#100ms;
	END_VAR

	VAR_OUTPUT
		XQ :	BOOL;
	END_VAR

	VAR
		tonRDMTimer :	TON;
		tof_xQ :	TOF;
		tRDMTime :	TIME;
		rRDMTime :	REAL;
		rdm_1 :	RDM_Block;
	END_VAR

	tonRDMTimer(IN:=Enable,PT:=tRDMTime);
	tof_xQ(IN := tonRDMTimer.Q,PT:=TP_Q);
	XQ := tof_xq.Q;
	IF tonRDMTimer.Q THEN
		xQ := TRUE ;
		rdm_1(last:=rRDMTime);
		rRDMTime:= rdm_1.RDM;

		tRDMTime := REAL_TO_TIME2(rRDMTime * TIME_TO_REAL1(Max_Time_ms - Min_Time_ms) + TIME_TO_REAL1(Min_Time_ms));
		tonRDMTimer (IN:=FALSE);
	END_IF;

END_FUNCTION_BLOCK

PROGRAM program0
  VAR
	ENABLE :	BOOL := TRUE;
	MIN_TIME_MS :	TIME := t#1s;
	MAX_TIME_MS :	TIME := t#1.2s;
	TP_Q :	TIME := t#100ms;
	XQ :	BOOL;
	func_block : GEN_RDT_Block;
  END_VAR
	func_block.ENABLE  :=ENABLE;
	func_block.MIN_TIME_MS  :=MIN_TIME_MS;
	func_block.MAX_TIME_MS  :=MAX_TIME_MS;
	func_block.TP_Q  :=TP_Q;
	func_block();
	XQ := func_block.XQ;
END_PROGRAM

CONFIGURATION Config0
	VAR_GLOBAL
		PLC_TICKS_PER_SEC :	INT;
		PLC_SYS_TICK_CNT :	DINT;
	END_VAR
	RESOURCE Res0 ON PLC
		TASK task0(INTERVAL := T#20ms,PRIORITY := 0);
		PROGRAM instance0 WITH task0 : program0;
	END_RESOURCE
END_CONFIGURATION

(* ---- 696-FT_PIDW.ST ---- *)
FUNCTION _REAL_TO_UDINT:UDINT
  VAR_INPUT
    X :	REAL;
  END_VAR

  IF REAL_TO_UDINT(0.5) = UDINT#1 THEN
    _REAL_TO_UDINT := REAL_TO_UDINT(x);
  ELSIF X > 0.0 THEN
    _REAL_TO_UDINT := REAL_TO_UDINT(x+0.5);
  ELSIF X < 0.0 THEN
    _REAL_TO_UDINT := REAL_TO_UDINT(x-0.5);
  ELSE
    _REAL_TO_UDINT := UDINT#0;
  END_IF;
END_FUNCTION

FUNCTION REAL_TO_TIME2:TIME
	VAR_INPUT
		IN :	REAL;
	END_VAR

	REAL_TO_TIME2 := DINT_TO_TIME(UDINT_TO_DINT(_REAL_TO_UDINT(IN)));
END_FUNCTION

FUNCTION_BLOCK T_PLC_US_Block
	VAR_OUTPUT
		T_PLC_US :	UDINT;
	END_VAR

	VAR_EXTERNAL
		PLC_TICKS_PER_SEC :	INT;
		PLC_SYS_TICK_CNT :	DINT;
	END_VAR

	VAR
		debug :	BOOL;
		N :	INT;
		Offset :	UDINT;
		temp :	DWORD := DWORD#1;
		mode :	BOOL;
		faktor :	UDINT;
		init :	BOOL;
		v_plc_ticks_per_sec :	UDINT;
		base :	UDINT := UDINT#1000000;
	END_VAR

	IF init = FALSE THEN
		v_plc_ticks_per_sec := INT_TO_UDINT(PLC_TICKS_PER_SEC);
		IF v_plc_ticks_per_sec = UDINT#1024 THEN
			faktor := UDINT#1000;
			mode := FALSE;
		ELSIF v_plc_ticks_per_sec > UDINT#0 THEN
			IF v_plc_ticks_per_sec <= base THEN
				faktor := base / v_plc_ticks_per_sec;
				mode := FALSE;
			ELSE
				faktor := v_plc_ticks_per_sec / base;
				mode := TRUE;
			END_IF;
		ELSE
			faktor := UDINT#1;
		END_IF;
		init := TRUE;
	END_IF;

	IF mode THEN
		T_PLC_US := DINT_TO_UDINT(PLC_SYS_TICK_CNT) / faktor;
	ELSE
		T_PLC_US := DINT_TO_UDINT(PLC_SYS_TICK_CNT) * faktor;
	END_IF;

	IF debug THEN
		T_PLC_US := (DWORD_TO_UDINT(SHL(UDINT_TO_DWORD(T_PLC_US),N) OR SHL(temp,N)) - UDINT#1) + Offset;
	END_IF;
END_FUNCTION_BLOCK

FUNCTION_BLOCK FT_DERIV
	VAR_INPUT
		IN :	REAL;
		K :	REAL := 1.0;
		RUN :	BOOL := TRUE;
	END_VAR

	VAR_OUTPUT
		OUT :	REAL;
	END_VAR

	VAR
		old :	REAL;
		tx :	UDINT;
		last :	UDINT;
		init :	BOOL;
		tc :	REAL;
		T_PLC_US :	T_PLC_US_Block;
	END_VAR

	T_PLC_US();
	tx:= T_PLC_US.T_PLC_US;
	tc := UDINT_TO_REAL(tx - last);

	IF NOT init THEN
		init := TRUE;
		old := in;
	ELSIF run AND tc > 0.0 THEN
		out := (in - old) / tc * 1000000.0 * K;
		old := in;
	ELSE
		out := 0.0;
	END_IF;

	last := tx;

	T_PLC_US();
	tx:= T_PLC_US.T_PLC_US;

	IF NOT init THEN
		init := TRUE;
	ELSIF run AND tx - last > UDINT#0 THEN
		out := (in - old) / UDINT_TO_REAL(tx - last) * 1000000.0 * K;
	ELSE
		out := 0.0;
	END_IF;
	old := in;
	last := tx;
END_FUNCTION_BLOCK
FUNCTION_BLOCK T_PLC_MS_block
	VAR_OUTPUT
		T_PLC_MS :	UDINT;
	END_VAR

	VAR_EXTERNAL
		PLC_TICKS_PER_SEC :	INT;
		PLC_SYS_TICK_CNT :	DINT;
	END_VAR

	VAR
		debug :	BOOL;(*Debug-Mode ON / OFF*)
		N :	INT;(*Debug-Faktor*)
		Offset :	UDINT;(*Debug-Offset*)
		temp :	DWORD := DWORD#1;(*Debug-Offset*)
		mode :	BOOL;(*modus*)
		faktor :	UDINT;(*Systemtakt-Faktor*)
		init :	BOOL;
		v_plc_ticks_per_sec :	UDINT;
		base :	UDINT := UDINT#1000;
	END_VAR

	IF init = FALSE THEN
		v_plc_ticks_per_sec := INT_TO_UDINT(PLC_TICKS_PER_SEC);
		IF v_plc_ticks_per_sec = UDINT#1024 THEN
			faktor := UDINT#1;
			mode := FALSE;
		ELSIF v_plc_ticks_per_sec > UDINT#0 THEN
			IF v_plc_ticks_per_sec <= base THEN
				faktor := base / v_plc_ticks_per_sec;
				mode := FALSE;
			ELSE
				faktor := v_plc_ticks_per_sec / base;
				mode := TRUE;
			END_IF;
		ELSE
			faktor := UDINT#1;
		END_IF;
		init := TRUE;
	END_IF;

	IF mode THEN
		T_PLC_MS := DINT_TO_UDINT(PLC_SYS_TICK_CNT) / faktor;
	ELSE
		T_PLC_MS := DINT_TO_UDINT(PLC_SYS_TICK_CNT) * faktor;
	END_IF;

	IF debug THEN
		T_PLC_MS := (DWORD_TO_UDINT(SHL(UDINT_TO_DWORD(T_PLC_MS),N) OR SHL(temp,N)) - UDINT#1) + Offset;
	END_IF;
END_FUNCTION_BLOCK

FUNCTION_BLOCK INTEGRATE

	VAR_INPUT
		E :	BOOL := TRUE;
		X :	REAL;
		K :	REAL := 1.0;
	END_VAR

	VAR_IN_OUT
		Y :	REAL;
	END_VAR

	VAR
		X_last :	REAL;
		init :	BOOL;
		T_PLC_MS :	T_PLC_MS_block;
		last :	UDINT;
		tx :	UDINT;
	END_VAR

	T_PLC_MS();
	tx:= T_PLC_MS.T_PLC_MS;

	IF NOT init THEN
		init := TRUE;
		X_last := X;
	ELSIF E THEN
		Y := (X + X_LAST) * 0.5E-3 * UDINT_TO_REAL(tx-last) * K + Y;
		X_last := X;
	END_IF;
	last := tx;

END_FUNCTION_BLOCK

FUNCTION_BLOCK FT_PIDW

	VAR_INPUT
		IN :	REAL;
		KP :	REAL := 1.0;
		TN :	REAL := 1.0;
		TV :	REAL := 1.0;
		LIM_L :	REAL := -1.0E38;
		LIM_H :	REAL := 1.0E38;
		RST :	BOOL := FALSE;
	END_VAR

	VAR_OUTPUT
		Y :	REAL;
		LIM :	BOOL;
	END_VAR

	VAR
		integ :	INTEGRATE;
		diff :	FT_DERIV;
		YI :	REAL;
	END_VAR

	IF tn = 0.0 OR rst THEN
		integ(E := FALSE, Y := YI);
		YI := integ.Y;
		YI := 0.0;
	ELSE
		integ(X := IN, K := 1.0 / TN, E := NOT LIM, Y := YI);
		YI := integ.Y;
	END_IF;

	(* add up integrator and linear part *)
	Y := KP * (IN + YI);

	(* run differentiator *)
	diff(IN := IN, K := TV);

	(* set lim before differentiator is added to stop integrator if necessary *)
	IF Y > LIM_L AND Y < LIM_H THEN
		LIM := FALSE;
	ELSE
		LIM := TRUE;
	END_IF;

	Y := LIMIT(LIM_L, Y + KP * diff.out, LIM_H);

END_FUNCTION_BLOCK

PROGRAM program0
	VAR
		IN :	REAL;
		KP :	REAL := 1.0;
		TN :	REAL := 1.0;
		TV :	REAL := 1.0;
		LIM_L :	REAL := -1.0E38;
		LIM_H :	REAL := 1.0E38;
		RST :	BOOL := FALSE;

		Y :	REAL;
		LIM :	BOOL;

		func_block : FT_PIDW;
	END_VAR
	func_block.IN := IN;
	func_block.KP := KP;
	func_block.TN := TN;
	func_block.TV := TV;
	func_block.LIM_L := LIM_L;
	func_block.LIM_H := LIM_H;
	func_block.RST := RST;

	func_block();
	Y := func_block.Y;
	LIM := func_block.LIM;
END_PROGRAM

CONFIGURATION Config0

	VAR_GLOBAL
		PLC_TICKS_PER_SEC :	INT;
		PLC_SYS_TICK_CNT :	DINT;
	END_VAR

	RESOURCE Res0 ON PLC
		TASK task0(INTERVAL := T#20ms,PRIORITY := 0);
		PROGRAM instance0 WITH task0 : program0;
	END_RESOURCE

END_CONFIGURATION

(* ---- 697-FT_PID.ST ---- *)
FUNCTION_BLOCK T_PLC_US_Block
	VAR_OUTPUT
		T_PLC_US :	UDINT;
	END_VAR

	VAR_EXTERNAL
		PLC_TICKS_PER_SEC :	INT;
		PLC_SYS_TICK_CNT :	DINT;
	END_VAR

	VAR
		debug :	BOOL;
		N :	INT;
		Offset :	UDINT;
		temp :	DWORD := DWORD#1;
		mode :	BOOL;
		faktor :	UDINT;
		init :	BOOL;
		v_plc_ticks_per_sec :	UDINT;
		base :	UDINT := UDINT#1000000;
	END_VAR

	IF init = FALSE THEN
		v_plc_ticks_per_sec := INT_TO_UDINT(PLC_TICKS_PER_SEC);
		IF v_plc_ticks_per_sec = UDINT#1024 THEN
			faktor := UDINT#1000;
			mode := FALSE;
		ELSIF v_plc_ticks_per_sec > UDINT#0 THEN
			IF v_plc_ticks_per_sec <= base THEN
				faktor := base / v_plc_ticks_per_sec;
				mode := FALSE;
			ELSE
				faktor := v_plc_ticks_per_sec / base;
				mode := TRUE;
			END_IF;
		ELSE
			faktor := UDINT#1;
		END_IF;
		init := TRUE;
	END_IF;

	IF mode THEN
		T_PLC_US := DINT_TO_UDINT(PLC_SYS_TICK_CNT) / faktor;
	ELSE
		T_PLC_US := DINT_TO_UDINT(PLC_SYS_TICK_CNT) * faktor;
	END_IF;

	IF debug THEN
		T_PLC_US := (DWORD_TO_UDINT(SHL(UDINT_TO_DWORD(T_PLC_US),N) OR SHL(temp,N)) - UDINT#1) + Offset;
	END_IF;
END_FUNCTION_BLOCK

FUNCTION_BLOCK T_PLC_MS_block
	VAR_OUTPUT
		T_PLC_MS :	UDINT;
	END_VAR

	VAR_EXTERNAL
		PLC_TICKS_PER_SEC :	INT;
		PLC_SYS_TICK_CNT :	DINT;
	END_VAR

	VAR
		debug :	BOOL;(*Debug-Mode ON / OFF*)
		N :	INT;(*Debug-Faktor*)
		Offset :	UDINT;(*Debug-Offset*)
		temp :	DWORD := DWORD#1;(*Debug-Offset*)
		mode :	BOOL;(*modus*)
		faktor :	UDINT;(*Systemtakt-Faktor*)
		init :	BOOL;
		v_plc_ticks_per_sec :	UDINT;
		base :	UDINT := UDINT#1000;
	END_VAR

	IF init = FALSE THEN
		v_plc_ticks_per_sec := INT_TO_UDINT(PLC_TICKS_PER_SEC);
		IF v_plc_ticks_per_sec = UDINT#1024 THEN
			faktor := UDINT#1;
			mode := FALSE;
		ELSIF v_plc_ticks_per_sec > UDINT#0 THEN
			IF v_plc_ticks_per_sec <= base THEN
				faktor := base / v_plc_ticks_per_sec;
				mode := FALSE;
			ELSE
				faktor := v_plc_ticks_per_sec / base;
				mode := TRUE;
			END_IF;
		ELSE
			faktor := UDINT#1;
		END_IF;
		init := TRUE;
	END_IF;

	IF mode THEN
		T_PLC_MS := DINT_TO_UDINT(PLC_SYS_TICK_CNT) / faktor;
	ELSE
		T_PLC_MS := DINT_TO_UDINT(PLC_SYS_TICK_CNT) * faktor;
	END_IF;

	IF debug THEN
		T_PLC_MS := (DWORD_TO_UDINT(SHL(UDINT_TO_DWORD(T_PLC_MS),N) OR SHL(temp,N)) - UDINT#1) + Offset;
	END_IF;
END_FUNCTION_BLOCK

FUNCTION_BLOCK INTEGRATE

	VAR_INPUT
		E :	BOOL := TRUE;
		X :	REAL;
		K :	REAL := 1.0;
	END_VAR

	VAR_IN_OUT
		Y :	REAL;
	END_VAR

	VAR
		X_last :	REAL;
		init :	BOOL;
		T_PLC_MS :	T_PLC_MS_block;
		last :	UDINT;
		tx :	UDINT;
	END_VAR

	T_PLC_MS();
	tx:= T_PLC_MS.T_PLC_MS;

	IF NOT init THEN
		init := TRUE;
		X_last := X;
	ELSIF E THEN
		Y := (X + X_LAST) * 0.5E-3 * UDINT_TO_REAL(tx-last) * K + Y;
		X_last := X;
	END_IF;
	last := tx;

END_FUNCTION_BLOCK

FUNCTION_BLOCK FT_INT_Block

	VAR_INPUT
		IN :	REAL;
		K :	REAL := 1.0;
		RUN :	BOOL := TRUE;
		RST :	BOOL;
		OUT_MIN :	REAL := REAL#-1.0E-37;
		OUT_MAX :	REAL := REAL#1.0E37;
	END_VAR

	VAR_OUTPUT
		OUT :	REAL;
		LIM :	BOOL;
	END_VAR

	VAR
		INTEG :	INTEGRATE;
	END_VAR

	IF rst THEN
		out := 0.0;
	ELSE
		integ(X := IN, E := RUN, K := K, Y := out);
		out := integ.Y;
	END_IF;

	(* limit the outputs *)
	IF out >= OUT_MAX THEN
		out := out_max;
		LIM := TRUE;
	ELSIF out <= out_min THEN
		out := out_min;
		lim := TRUE;
	ELSE
		lim := FALSE;
	END_IF;

END_FUNCTION_BLOCK

FUNCTION_BLOCK FT_DERIV
	VAR_INPUT
		IN :	REAL;
		K :	REAL := 1.0;
		RUN :	BOOL := TRUE;
	END_VAR

	VAR_OUTPUT
		OUT :	REAL;
	END_VAR

	VAR
		old :	REAL;
		tx :	UDINT;
		last :	UDINT;
		init :	BOOL;
		tc :	REAL;
		T_PLC_US :	T_PLC_US_Block;
	END_VAR

	T_PLC_US();
	tx:= T_PLC_US.T_PLC_US;
	tc := UDINT_TO_REAL(tx - last);

	IF NOT init THEN
		init := TRUE;
		old := in;
	ELSIF run AND tc > 0.0 THEN
		out := (in - old) / tc * 1000000.0 * K;
		old := in;
	ELSE
		out := 0.0;
	END_IF;

	last := tx;

	T_PLC_US();
	tx:= T_PLC_US.T_PLC_US;

	IF NOT init THEN
		init := TRUE;
	ELSIF run AND tx - last > UDINT#0 THEN
		out := (in - old) / UDINT_TO_REAL(tx - last) * 1000000.0 * K;
	ELSE
		out := 0.0;
	END_IF;
	old := in;
	last := tx;
END_FUNCTION_BLOCK

FUNCTION_BLOCK FT_PID

	VAR_INPUT
		IN :	REAL;
		KP :	REAL := 1.0;
		TN :	REAL := 1.0;
		TV :	REAL := 1.0;
		ILIM_L :	REAL := -1.0E38;
		ILIM_H :	REAL := 1.0E38;
		IEN :	BOOL := TRUE;
		RST :	BOOL := FALSE;
	END_VAR

	VAR_OUTPUT
		Y :	REAL;
		LIM :	BOOL;
	END_VAR

	VAR
		integ :	FT_INT_Block;
		diff :	FT_DERIV;
	END_VAR

	IF TN > 0.0 THEN
		integ(IN := IN, K := 1.0 / TN, RUN := IEN, RST := RST, OUT_MIN := ILIM_L, OUT_MAX := ILIM_H);
	ELSE
		integ(RST := FALSE);
	END_IF;

	(* run differentiator *)
	diff(IN := IN, K := TV);

	(* combine both values *)
	Y := KP * (integ.Out + diff.out + IN);

	(* check if integrator has reached its limits and set overflow *)
	LIM := integ.LIM;

END_FUNCTION_BLOCK

PROGRAM program0
	VAR
		IN :	REAL;
		KP :	REAL := 1.0;
		TN :	REAL := 1.0;
		TV :	REAL := 1.0;
		ILIM_L :	REAL := -1.0E38;
		ILIM_H :	REAL := 1.0E38;
		IEN :	BOOL := TRUE;
		RST :	BOOL := FALSE;

		Y :	REAL;
		LIM :	BOOL;

		func_block : FT_PID;
	END_VAR
	func_block.IN :=IN;
	func_block.KP :=KP;
	func_block.TN :=TN;
	func_block.TV :=TV;
	func_block.ILIM_L :=ILIM_L;
	func_block.ILIM_H :=ILIM_H;
	func_block.IEN :=IEN;
	func_block.RST :=RST;

	func_block();
	Y := func_block.Y;
	LIM := func_block.LIM;
END_PROGRAM

CONFIGURATION Config0

	VAR_GLOBAL
		PLC_TICKS_PER_SEC :	INT;
		PLC_SYS_TICK_CNT :	DINT;
	END_VAR

	RESOURCE Res0 ON PLC
		TASK task0(INTERVAL := T#20ms,PRIORITY := 0);
		PROGRAM instance0 WITH task0 : program0;
	END_RESOURCE

END_CONFIGURATION

(* ---- 698-PARSET.ST ---- *)
TYPE
	oscat_parset_X              : ARRAY [1..4]    OF REAL;
	oscat_parset                : ARRAY [0..3]    OF oscat_parset_X := [0,0,0,0];
END_TYPE

FUNCTION TIME_TO_UDINT2:UDINT
	VAR_INPUT
		X :	TIME;
	END_VAR

	TIME_TO_UDINT2 := DINT_TO_UDINT(TIME_TO_DINT(X));
END_FUNCTION

FUNCTION _BYTE_TO_INT:INT
	VAR_INPUT
		IN :	BYTE;
	END_VAR

	_BYTE_TO_INT := USINT_TO_INT(BYTE_TO_USINT(IN));
END_FUNCTION

FUNCTION BIT_OF_DWORD : BOOL
  VAR_INPUT
    IN : DWORD;
    N : INT;
  END_VAR

  BIT_OF_DWORD := (SHR(in,N) AND 16#00000001) > 0;
  (* from OSCAT library; www.oscat.de  *)
END_FUNCTION

FUNCTION BIT_LOAD_B:BYTE
	VAR_INPUT
		IN :	BYTE;
		VAL :	BOOL;
		POS :	INT;
	END_VAR

	IF VAL THEN
		BIT_LOAD_B := in OR SHL(BYTE#1,pos);
	ELSE
		BIT_LOAD_B := in AND (NOT SHL(BYTE#1,pos));
	END_IF;
END_FUNCTION

FUNCTION_BLOCK T_PLC_MS_block
	VAR_OUTPUT
		T_PLC_MS :	UDINT;
	END_VAR

	VAR_EXTERNAL
		PLC_TICKS_PER_SEC :	INT;
		PLC_SYS_TICK_CNT :	DINT;
	END_VAR

	VAR
		debug :	BOOL;(*Debug-Mode ON / OFF*)
		N :	INT;(*Debug-Faktor*)
		Offset :	UDINT;(*Debug-Offset*)
		temp :	DWORD := DWORD#1;(*Debug-Offset*)
		mode :	BOOL;(*modus*)
		faktor :	UDINT;(*Systemtakt-Faktor*)
		init :	BOOL;
		v_plc_ticks_per_sec :	UDINT;
		base :	UDINT := UDINT#1000;
	END_VAR

	IF init = FALSE THEN
		v_plc_ticks_per_sec := INT_TO_UDINT(PLC_TICKS_PER_SEC);
		IF v_plc_ticks_per_sec = UDINT#1024 THEN
			faktor := UDINT#1;
			mode := FALSE;
		ELSIF v_plc_ticks_per_sec > UDINT#0 THEN
			IF v_plc_ticks_per_sec <= base THEN
				faktor := base / v_plc_ticks_per_sec;
				mode := FALSE;
			ELSE
				faktor := v_plc_ticks_per_sec / base;
				mode := TRUE;
			END_IF;
		ELSE
			faktor := UDINT#1;
		END_IF;
		init := TRUE;
	END_IF;

	IF mode THEN
		T_PLC_MS := DINT_TO_UDINT(PLC_SYS_TICK_CNT) / faktor;
	ELSE
		T_PLC_MS := DINT_TO_UDINT(PLC_SYS_TICK_CNT) * faktor;
	END_IF;

	IF debug THEN
		T_PLC_MS := (DWORD_TO_UDINT(SHL(UDINT_TO_DWORD(T_PLC_MS),N) OR SHL(temp,N)) - UDINT#1) + Offset;
	END_IF;
END_FUNCTION_BLOCK

FUNCTION_BLOCK PARSET_Block

	VAR_INPUT
		A0 :	BOOL;
		A1 :	BOOL;
		X01 :	REAL;
		X02 :	REAL;
		X03 :	REAL;
		X04 :	REAL;
		X11 :	REAL;
		X12 :	REAL;
		X13 :	REAL;
		X14 :	REAL;
		X21 :	REAL;
		X22 :	REAL;
		X23 :	REAL;
		X24 :	REAL;
		X31 :	REAL;
		X32 :	REAL;
		X33 :	REAL;
		X34 :	REAL;
		TC :	TIME;
	END_VAR

	VAR_OUTPUT
		P1 :	REAL;
		P2 :	REAL;
		P3 :	REAL;
		P4 :	REAL;
	END_VAR

	VAR
		X :	oscat_parset;
		S1 :	REAL;
		S2 :	REAL;
		S3 :	REAL;
		S4 :	REAL;
		tx :	UDINT;
		last :	UDINT;
		start :	BOOL;
		set :	BYTE;
		set2 :	INT;
		init :	BOOL;
		T_PLC_MS :	T_PLC_MS_Block;
	END_VAR

	(*@KEY@: WORKSHEET
	NAME: PARSET
	IEC_LANGUAGE: ST
	*)
	(* read system_time *)
	T_PLC_MS();
	tx:= T_PLC_MS.T_PLC_MS;

	(* init sequence *)
	IF NOT init THEN
		set:=BIT_LOAD_B(set,NOT A0,0); (* set.X0 := NOT A0; *)
		init := TRUE;
		X[0][1] := X01;
		X[0][2] := X02;
		X[0][3] := X03;
		X[0][4] := X04;
		X[1][1] := X11;
		X[1][2] := X12;
		X[1][3] := X13;
		X[1][4] := X14;
		X[2][1] := X21;
		X[2][2] := X22;
		X[2][3] := X23;
		X[2][4] := X24;
		X[3][1] := X31;
		X[3][2] := X32;
		X[3][3] := X33;
		X[3][4] := X34;
		P1 := X01;
		P2 := X02;
		P3 := X03;
		P4 := X04;
	END_IF;

	(* check for input change *)
	IF (A0 XOR BIT_OF_DWORD(BYTE_TO_DWORD(set),0)) OR (A1 XOR BIT_OF_DWORD(BYTE_TO_DWORD(set),1)) THEN  (* set.X0  ,  set.X1 *)
		(* a new set is selected *)
		set := BIT_LOAD_B(set,A0,0); (* set.X0 := A0; *)
		set := BIT_LOAD_B(set,A1,1); (* set.X1 := A1; *)

		IF tc > t#0s THEN
			start := TRUE;
			last := tx;
			(* save the step speed for the output changes in S *)
			set2 := _BYTE_TO_INT(set);
			S1 := (X[set2][1] - P1)/TIME_TO_REAL(tc);
			S2 := (X[set2][2] - P2)/TIME_TO_REAL(tc);
			S3 := (X[set2][3] - P3)/TIME_TO_REAL(tc);
			S4 := (X[set2][4] - P4)/TIME_TO_REAL(tc);
		END_IF;
	ELSIF start AND tx - last < TIME_TO_UDINT2(tc) THEN
		(* ramp the outputs to the new value *)
		set2 := _BYTE_TO_INT(set);
		P1 := X[set2][1] - S1*(TIME_TO_REAL(Tc) - UDINT_TO_REAL(tx + last));
		P2 := X[set2][2] - S2*(TIME_TO_REAL(Tc) - UDINT_TO_REAL(tx + last));
		P3 := X[set2][3] - S3*(TIME_TO_REAL(Tc) - UDINT_TO_REAL(tx + last));
		P4 := X[set2][4] - S4*(TIME_TO_REAL(Tc) - UDINT_TO_REAL(tx + last));
	ELSE
		(* make sure outputs match the correct set values *)
		set2 := _BYTE_TO_INT(set);
		start := FALSE;
		P1 := X[set2][1];
		P2 := X[set2][2];
		P3 := X[set2][3];
		P4 := X[set2][4];
	END_IF;

END_FUNCTION_BLOCK

PROGRAM program0

	VAR
		A0 :	BOOL;
		A1 :	BOOL;
		X01 :	REAL;
		X02 :	REAL;
		X03 :	REAL;
		X04 :	REAL;
		X11 :	REAL;
		X12 :	REAL;
		X13 :	REAL;
		X14 :	REAL;
		X21 :	REAL;
		X22 :	REAL;
		X23 :	REAL;
		X24 :	REAL;
		X31 :	REAL;
		X32 :	REAL;
		X33 :	REAL;
		X34 :	REAL;
		TC :	TIME;

		P1 :	REAL;
		P2 :	REAL;
		P3 :	REAL;
		P4 :	REAL;
		func_block : PARSET_Block;
  	END_VAR
	func_block.A0 := A0;
	func_block.A1 := A1;
	func_block.X01 := X01;
	func_block.X02 := X02;
	func_block.X03 := X03;
	func_block.X04 := X04;
	func_block.X11 := X11;
	func_block.X12 := X12;
	func_block.X13 := X13;
	func_block.X14 := X14;
	func_block.X21 := X21;
	func_block.X22 := X22;
	func_block.X23 := X23;
	func_block.X24 := X24;
	func_block.X31 := X31;
	func_block.X32 := X32;
	func_block.X33 := X33;
	func_block.X34 := X34;
	func_block.TC := TC;
	func_block();
	P1 := func_block.P1;
	P2 := func_block.P2;
	P3 := func_block.P3;
	P4 := func_block.P4;

END_PROGRAM

CONFIGURATION Config0

	VAR_GLOBAL
		PLC_TICKS_PER_SEC :	INT;
		PLC_SYS_TICK_CNT :	DINT;
	END_VAR

  	RESOURCE Res0 ON PLC
    	TASK task0(INTERVAL := T#20ms,PRIORITY := 0);
    	PROGRAM instance0 WITH task0 : program0;
  	END_RESOURCE

END_CONFIGURATION

(* ---- 699-ESR_MON_R4.ST ---- *)
TYPE
	oscat_esr_collect_data      : ARRAY [0..7]    OF BYTE;
END_TYPE

TYPE oscat_esr_data :
  STRUCT
	typ    : BYTE;
	adress : STRING;
	DS     : UDINT;
	TS     : TIME;
	data   : oscat_esr_collect_data;
  END_STRUCT;
END_TYPE

TYPE
  oscat_ESR_3                : ARRAY [0..3] OF oscat_esr_data;
  oscat_ESR_31               : ARRAY [0..31] OF oscat_esr_data;
END_TYPE

FUNCTION_BLOCK REAL_TO_DW_Block
  VAR_INPUT
    X :	REAL;
  END_VAR

  VAR_OUTPUT
    REAL_TO_DW :	DWORD;
  END_VAR

  VAR
    REAL_TO_BUF :	REAL_TO_BUF;
    i :	INT;
  END_VAR

  FOR I := 0 TO 1 DO
    REAL_TO_BUF.REQ        := I > 0;
    REAL_TO_BUF.BUF_FORMAT := FALSE;
    REAL_TO_BUF.BUF_OFFS   := DINT#0;
    REAL_TO_BUF.BUF_CNT    := DINT#4;
    REAL_TO_BUF.SRC        := X;
    REAL_TO_BUF.BUFFER     := REAL_TO_DW;
    REAL_TO_BUF();
    X          := REAL_TO_BUF.SRC;
    REAL_TO_DW := REAL_TO_BUF.BUFFER;
  END_FOR;
END_FUNCTION_BLOCK

FUNCTION_BLOCK T_PLC_MS_block

	VAR_OUTPUT
		T_PLC_MS :	UDINT;
	END_VAR

	VAR_EXTERNAL
		PLC_TICKS_PER_SEC :	INT;
		PLC_SYS_TICK_CNT :	DINT;
	END_VAR

	VAR
		debug :	BOOL;(*Debug-Mode ON / OFF*)
		N :	INT;(*Debug-Faktor*)
		Offset :	UDINT;(*Debug-Offset*)
		temp :	DWORD := DWORD#1;(*Debug-Offset*)
		mode :	BOOL;(*modus*)
		faktor :	UDINT;(*Systemtakt-Faktor*)
		init :	BOOL;
		v_plc_ticks_per_sec :	UDINT;
		base :	UDINT := UDINT#1000;
	END_VAR

	IF init = FALSE THEN
		v_plc_ticks_per_sec := INT_TO_UDINT(PLC_TICKS_PER_SEC);
		IF v_plc_ticks_per_sec = UDINT#1024 THEN
			faktor := UDINT#1;
			mode := FALSE;
		ELSIF v_plc_ticks_per_sec > UDINT#0 THEN
			IF v_plc_ticks_per_sec <= base THEN
				faktor := base / v_plc_ticks_per_sec;
				mode := FALSE;
			ELSE
				faktor := v_plc_ticks_per_sec / base;
				mode := TRUE;
			END_IF;
		ELSE
			faktor := UDINT#1;
		END_IF;
		init := TRUE;
	END_IF;

	IF mode THEN
		T_PLC_MS := DINT_TO_UDINT(PLC_SYS_TICK_CNT) / faktor;
	ELSE
		T_PLC_MS := DINT_TO_UDINT(PLC_SYS_TICK_CNT) * faktor;
	END_IF;

	IF debug THEN
		T_PLC_MS := (DWORD_TO_UDINT(SHL(UDINT_TO_DWORD(T_PLC_MS),N) OR SHL(temp,N)) - UDINT#1) + Offset;
	END_IF;

END_FUNCTION_BLOCK

FUNCTION_BLOCK ESR_MON_R4
	VAR_INPUT
		R0 :	REAL;
		A0 :	STRING;
		S0 :	REAL;
		R1 :	REAL;
		A1 :	STRING;
		S1 :	REAL;
		R2 :	REAL;
		A2 :	STRING;
		S2 :	REAL;
		R3 :	REAL;
		A3 :	STRING;
		S3 :	REAL;
		DT_IN :	UDINT;
	END_VAR

	VAR_IN_OUT
		ESR_OUT :	oscat_ESR_3;
	END_VAR

	VAR_OUTPUT
		ESR_FLAG :	BOOL;
	END_VAR

	VAR
		x0 :	REAL;
		x1 :	REAL;
		x2 :	REAL;
		x3 :	REAL;
		tx :	TIME;
		cnt :	INT;
		T_PLC_MS :	T_PLC_MS_block;
		REAL_TO_DW :	REAL_TO_DW_Block;
		tmp :	DWORD;
	END_VAR

	T_PLC_MS();
	tx:= UDINT_TO_TIME(T_PLC_MS.T_PLC_MS);

	ESR_Flag := FALSE;
	esr_out[3].typ := BYTE#0;
	esr_out[2].typ := BYTE#0;
	esr_out[1].typ := BYTE#0;
	esr_out[0].typ := BYTE#0;
	cnt := 0;

	IF differ(R0, X0, S0) THEN
		REAL_TO_DW(X:=R0);
		tmp := REAL_TO_DW.REAL_TO_DW;

		esr_out[cnt].typ := BYTE#20;
		esr_out[cnt].adress := a0;
		esr_out[cnt].DS := DT_in;
		esr_out[cnt].TS := TX;
		esr_out[cnt].data[0] := Byte_of_Dword(tmp,BYTE#0);
		esr_out[cnt].data[1] := Byte_of_Dword(tmp,BYTE#1);
		esr_out[cnt].data[2] := Byte_of_Dword(tmp,BYTE#2);
		esr_out[cnt].data[3] := Byte_of_Dword(tmp,BYTE#3);
		X0 := R0;
		cnt := cnt + 1;
		esr_flag := TRUE;
	END_IF;
	IF differ(R1, X1, S1) THEN
		REAL_TO_DW(X:=R1);
		tmp := REAL_TO_DW.REAL_TO_DW;

		esr_out[cnt].typ := BYTE#20;
		esr_out[cnt].adress := a1;
		esr_out[cnt].DS := DT_in;
		esr_out[cnt].TS := TX;
		esr_out[cnt].data[0] := Byte_of_Dword(tmp,BYTE#0);
		esr_out[cnt].data[1] := Byte_of_Dword(tmp,BYTE#1);
		esr_out[cnt].data[2] := Byte_of_Dword(tmp,BYTE#2);
		esr_out[cnt].data[3] := Byte_of_Dword(tmp,BYTE#3);
		X1 := R1;
		cnt := cnt + 1;
		esr_flag := TRUE;
	END_IF;
	IF differ(R2, X2, S2) THEN
		REAL_TO_DW(X:=R2);
		tmp := REAL_TO_DW.REAL_TO_DW;

		esr_out[cnt].typ := BYTE#20;
		esr_out[cnt].adress := a2;
		esr_out[cnt].DS := DT_in;
		esr_out[cnt].TS := TX;
		esr_out[cnt].data[0] := Byte_of_Dword(tmp,BYTE#0);
		esr_out[cnt].data[1] := Byte_of_Dword(tmp,BYTE#1);
		esr_out[cnt].data[2] := Byte_of_Dword(tmp,BYTE#2);
		esr_out[cnt].data[3] := Byte_of_Dword(tmp,BYTE#3);
		X2 := R2;
		cnt := cnt + 1;
		esr_flag := TRUE;
	END_IF;
	IF differ(R3, X3, S3) THEN
		REAL_TO_DW(X:=R2);
		tmp := REAL_TO_DW.REAL_TO_DW;

		esr_out[cnt].typ := BYTE#20;
		esr_out[cnt].adress := a3;
		esr_out[cnt].DS := DT_in;
		esr_out[cnt].TS := TX;
		esr_out[cnt].data[0] := Byte_of_Dword(tmp,BYTE#0);
		esr_out[cnt].data[1] := Byte_of_Dword(tmp,BYTE#1);
		esr_out[cnt].data[2] := Byte_of_Dword(tmp,BYTE#2);
		esr_out[cnt].data[3] := Byte_of_Dword(tmp,BYTE#3);
		X3 := R3;
		cnt := cnt + 1;
		esr_flag := TRUE;
	END_IF;
END_FUNCTION_BLOCK

PROGRAM program0

	VAR
	VAR_INPUT
		R0 :	REAL;
		A0 :	STRING;
		S0 :	REAL;
		R1 :	REAL;
		A1 :	STRING;
		S1 :	REAL;
		R2 :	REAL;
		A2 :	STRING;
		S2 :	REAL;
		R3 :	REAL;
		A3 :	STRING;
		S3 :	REAL;
		DT_IN :	UDINT;

		ESR_OUT :	oscat_ESR_3;

		ESR_FLAG :	BOOL;

		func_block : ESR_MON_R4;
  	END_VAR
	func_block.R0 := R0;
	func_block.A0 := A0;
	func_block.S0 := S0;
	func_block.R1 := R1;
	func_block.A1 := A1;
	func_block.S1 := S1;
	func_block.R2 := R2;
	func_block.A2 := A2;
	func_block.S2 := S2;
	func_block.R3 := R3;
	func_block.A3 := A3;
	func_block.S3 := S3;
	func_block.DT_IN := DT_IN;
	func_block.ESR_Out := ESR_Out;
	func_block();
	ESR_Out := func_block.ESR_Out;
	ESR_FLAG := func_block.ESR_FLAG;

END_PROGRAM

CONFIGURATION Config0

	VAR_GLOBAL
		PLC_TICKS_PER_SEC :	INT;
		PLC_SYS_TICK_CNT :	DINT;
	END_VAR

  	RESOURCE Res0 ON PLC
    	TASK task0(INTERVAL := T#20ms,PRIORITY := 0);
    	PROGRAM instance0 WITH task0 : program0;
  	END_RESOURCE

END_CONFIGURATION

(* ---- 700-MD5_STREAM.ST ---- *)
FUNCTION_BLOCK MD5_STREAM

	VAR_IN_OUT
		MODE :	INT;
		BUF :	oscat_aB0_63;
		MD5 :	oscat_aB0_15;
		SIZE :	UDINT;
	END_VAR

	VAR_OUTPUT
		POS :	UDINT;
	END_VAR

	VAR
		hash :	oscat_aDW0_3;
		a :	DWORD;
		b :	DWORD;
		c :	DWORD;
		d :	DWORD;
		end :	UDINT;
		block :	UDINT;
		x :	oscat_aDW0_15;
		pad_1 :	BOOL;
		n :	INT;
		n1 :	INT;
		n2 :	INT;
		n3 :	INT;
		n4 :	INT;
	END_VAR

	CASE MODE OF

	1:
		hash[0] := DWORD#16#67452301;
		hash[1] := DWORD#16#EFCDAB89;
		hash[2] := DWORD#16#98BADCFE;
		hash[3] := DWORD#16#10325476;

		block := DWORD_TO_UDINT(SHR_DWORD(UDINT_TO_DWORD(SIZE),6)) + BOOL_TO_UDINT((UDINT_TO_BYTE(SIZE) AND BYTE#16#3F) > BYTE#55);
		pad_1 := FALSE;
		POS := UDINT#0;
		End := SIZE;
		SIZE := MIN(UDINT#64,end);
		MODE := 2;

	2:
		FOR n := UDINT_TO_INT(SIZE) TO 63 DO
			BUF[n] := BYTE#0;
		END_FOR;

		IF SIZE < UDINT#64 AND NOT pad_1 THEN
			BUF[SIZE] := BYTE#2#1000_0000;
			pad_1 := TRUE;
		END_IF;

		POS := POS + SIZE;
		SIZE := MIN(UDINT#64,End - POS);

		n := 0;
		FOR n4 := 0 TO 15 DO
			n1 := n + 1;
			n2 := n + 2;
			n3 := n + 3;
			x[n4] := DWORD_OF_BYTE(BUF[n3],BUF[n2],BUF[n1],BUF[n]);
			n := n + 4;
		END_FOR;

		IF block = UDINT#0 THEN
			x[14] := SHL_DWORD(UDINT_TO_DWORD(End),3);
			MODE := 3;
		ELSE
			block := block - UDINT#1;
		END_IF;

		a := hash[0];
		b := hash[1];
		c := hash[2];
		d := hash[3];

		a := MD5_AUX(1, a, b, c, d, X[00], 07, DWORD#16#D76AA478);
		d := MD5_AUX(1, d, a, b, c, X[01], 12, DWORD#16#E8C7B756);
		c := MD5_AUX(1, c, d, a, b, X[02], 17, DWORD#16#242070DB);
		b := MD5_AUX(1, b, c, d, a, X[03], 22, DWORD#16#C1BDCEEE);
		a := MD5_AUX(1, a, b, c, d, X[04], 07, DWORD#16#F57C0FAF);
		d := MD5_AUX(1, d, a, b, c, X[05], 12, DWORD#16#4787C62A);
		c := MD5_AUX(1, c, d, a, b, X[06], 17, DWORD#16#A8304613);
		b := MD5_AUX(1, b, c, d, a, X[07], 22, DWORD#16#FD469501);
		a := MD5_AUX(1, a, b, c, d, X[08], 07, DWORD#16#698098D8);
		d := MD5_AUX(1, d, a, b, c, X[09], 12, DWORD#16#8B44F7AF);
		c := MD5_AUX(1, c, d, a, b, X[10], 17, DWORD#16#FFFF5BB1);
		b := MD5_AUX(1, b, c, d, a, X[11], 22, DWORD#16#895CD7BE);
		a := MD5_AUX(1, a, b, c, d, X[12], 07, DWORD#16#6B901122);
		d := MD5_AUX(1, d, a, b, c, X[13], 12, DWORD#16#FD987193);
		c := MD5_AUX(1, c, d, a, b, X[14], 17, DWORD#16#A679438E);
		b := MD5_AUX(1, b, c, d, a, X[15], 22, DWORD#16#49B40821);

		a := MD5_AUX(2, a, b, c, d, X[01], 05, DWORD#16#F61E2562);
		d := MD5_AUX(2, d, a, b, c, X[06], 09, DWORD#16#C040B340);
		c := MD5_AUX(2, c, d, a, b, X[11], 14, DWORD#16#265E5A51);
		b := MD5_AUX(2, b, c, d, a, X[00], 20, DWORD#16#E9B6C7AA);
		a := MD5_AUX(2, a, b, c, d, X[05], 05, DWORD#16#D62F105D);
		d := MD5_AUX(2, d, a, b, c, X[10], 09, DWORD#16#02441453);
		c := MD5_AUX(2, c, d, a, b, X[15], 14, DWORD#16#D8A1E681);
		b := MD5_AUX(2, b, c, d, a, X[04], 20, DWORD#16#E7D3FBC8);
		a := MD5_AUX(2, a, b, c, d, X[09], 05, DWORD#16#21E1CDE6);
		d := MD5_AUX(2, d, a, b, c, X[14], 09, DWORD#16#C33707D6);
		c := MD5_AUX(2, c, d, a, b, X[03], 14, DWORD#16#F4D50D87);
		b := MD5_AUX(2, b, c, d, a, X[08], 20, DWORD#16#455A14ED);
		a := MD5_AUX(2, a, b, c, d, X[13], 05, DWORD#16#A9E3E905);
		d := MD5_AUX(2, d, a, b, c, X[02], 09, DWORD#16#FCEFA3F8);
		c := MD5_AUX(2, c, d, a, b, X[07], 14, DWORD#16#676F02D9);
		b := MD5_AUX(2, b, c, d, a, X[12], 20, DWORD#16#8D2A4C8A);

		a := MD5_AUX(3, a, b, c, d, X[05], 04, DWORD#16#FFFA3942);
		d := MD5_AUX(3, d, a, b, c, X[08], 11, DWORD#16#8771F681);
		c := MD5_AUX(3, c, d, a, b, X[11], 16, DWORD#16#6D9D6122);
		b := MD5_AUX(3, b, c, d, a, X[14], 23, DWORD#16#FDE5380C);
		a := MD5_AUX(3, a, b, c, d, X[01], 04, DWORD#16#A4BEEA44);
		d := MD5_AUX(3, d, a, b, c, X[04], 11, DWORD#16#4BDECFA9);
		c := MD5_AUX(3, c, d, a, b, X[07], 16, DWORD#16#F6BB4B60);
		b := MD5_AUX(3, b, c, d, a, X[10], 23, DWORD#16#BEBFBC70);
		a := MD5_AUX(3, a, b, c, d, X[13], 04, DWORD#16#289B7EC6);
		d := MD5_AUX(3, d, a, b, c, X[00], 11, DWORD#16#EAA127FA);
		c := MD5_AUX(3, c, d, a, b, X[03], 16, DWORD#16#D4EF3085);
		b := MD5_AUX(3, b, c, d, a, X[06], 23, DWORD#16#04881D05);
		a := MD5_AUX(3, a, b, c, d, X[09], 04, DWORD#16#D9D4D039);
		d := MD5_AUX(3, d, a, b, c, X[12], 11, DWORD#16#E6DB99E5);
		c := MD5_AUX(3, c, d, a, b, X[15], 16, DWORD#16#1FA27CF8);
		b := MD5_AUX(3, b, c, d, a, X[02], 23, DWORD#16#C4AC5665);

		a := MD5_AUX(4, a, b, c, d, X[00], 06, DWORD#16#F4292244);
		d := MD5_AUX(4, d, a, b, c, X[07], 10, DWORD#16#432AFF97);
		c := MD5_AUX(4, c, d, a, b, X[14], 15, DWORD#16#AB9423A7);
		b := MD5_AUX(4, b, c, d, a, X[05], 21, DWORD#16#FC93A039);
		a := MD5_AUX(4, a, b, c, d, X[12], 06, DWORD#16#655B59C3);
		d := MD5_AUX(4, d, a, b, c, X[03], 10, DWORD#16#8F0CCC92);
		c := MD5_AUX(4, c, d, a, b, X[10], 15, DWORD#16#FFEFF47D);
		b := MD5_AUX(4, b, c, d, a, X[01], 21, DWORD#16#85845DD1);
		a := MD5_AUX(4, a, b, c, d, X[08], 06, DWORD#16#6FA87E4F);
		d := MD5_AUX(4, d, a, b, c, X[15], 10, DWORD#16#FE2CE6E0);
		c := MD5_AUX(4, c, d, a, b, X[06], 15, DWORD#16#A3014314);
		b := MD5_AUX(4, b, c, d, a, X[13], 21, DWORD#16#4E0811A1);
		a := MD5_AUX(4, a, b, c, d, X[04], 06, DWORD#16#F7537E82);
		d := MD5_AUX(4, d, a, b, c, X[11], 10, DWORD#16#BD3AF235);
		c := MD5_AUX(4, c, d, a, b, X[02], 15, DWORD#16#2AD7D2BB);
		b := MD5_AUX(4, b, c, d, a, X[09], 21, DWORD#16#EB86D391);

		hash[0] := UDINT_TO_DWORD(DWORD_TO_UDINT(hash[0]) + DWORD_TO_UDINT(a));
		hash[1] := UDINT_TO_DWORD(DWORD_TO_UDINT(hash[1]) + DWORD_TO_UDINT(b));
		hash[2] := UDINT_TO_DWORD(DWORD_TO_UDINT(hash[2]) + DWORD_TO_UDINT(c));
		hash[3] := UDINT_TO_DWORD(DWORD_TO_UDINT(hash[3]) + DWORD_TO_UDINT(d));

	END_CASE;

	IF MODE = 3 THEN
		n2 := 0;
		FOR n := 0 TO 3 DO
			FOR n1 := 0 TO 3 DO
				MD5[n2] := DWORD_TO_BYTE(hash[n]);
				hash[n] := ROR_DWORD(hash[n],8);
				n2 := n2 + 1;
			END_FOR;
		END_FOR;
	END_IF;

END_FUNCTION_BLOCK
